(* IEC 61131-3 sources: SortJet_MasterSPS_Aufbau.fbsproj/07_Auftragsverwaltung/BasisSchrittketten (part 2) *)

(* ---- Station_Austransport.fb.st ---- *)
(* METADATA
{
	"v3Meta": {
		"objectGuid": "ceff7ec0-8422-4f2f-902e-5124ad2e42bc"
	}
}
*)
FUNCTION_BLOCK Station_Austransport
VAR_INPUT

  // BOOLEAN
  bpReset                : BOOL;

  // WORD
  wStation               : WORD;
  wWand                  : WORD;

  // STRUKTUR
  Auftragsdaten          : Auftragsdaten_ST;

END_VAR
VAR_OUTPUT

  // BOOLEAN
  bpDone                 : BOOL;
  bpFehler               : BOOL;

END_VAR
VAR

  // BOOLEAN
  blStationQuittiertScheiben      : BOOL;
  blGegenstelleIstShuttle         : BOOL;

  // INT
  ilScheibenZuQuittieren          : INT;

  // WORD
  wlAustransportstation           : WORD;
  wlAustransportstationVorgaenger : WORD;

  // REFERENZ
  Gegenstelle                     : REFERENCE TO StationBasisParameter_ST;

  // STEPS
  steplSchritt           : STEPS_TE;

END_VAR
//-------------------------------------------------------------------------------------------------
// STEUERUNG AUSTRANSPORT
//-------------------------------------------------------------------------------------------------
IF Auftragsdaten.wAuftrag = eStation_Austransport THEN
  CASE steplSchritt OF
    // AUSTRANSPORT =================================
    STEP_0_E:
      (* Hinweis:
         - Ueberpruefung des Sicherheitskreises
      *)
      IF checkSafetyCircuitsNotBlocked(starrStationBasisParameter[wStation], eSKKomponente_Glastransport) THEN
        steplSchritt := STEP_10_E;
      END_IF

    // AUSTRANSPORT ==================================================
    STEP_10_E:
      // ---------------------------------------------------------------------------------------
      //  OPTIONALE - PRUEFUNG DER GLASDATEN
      //
      //  Hinweis:
      // - n/c
      // ---------------------------------------------------------------------------------------
      steplSchritt := STEP_20_E;

      IF NOT AuftragsdatenPruefen( wStation, wWand, Auftragsdaten) THEN
        steplSchritt := STEP_900_E;
      END_IF

    // AUSTRANSPORT =================================
    STEP_20_E:
      (* Hinweis:
         - Uebergabe der Quellstation [Sender] fuer den Austransport [Zum ueberpruefen des Zustandes der Station]
      *)
      wlAustransportstation := Auftragsdaten.wTransferstationsNr1;

      (* Hinweis:
         - Nach einem Systemcheck mit übergroßen Scheiben kann es sein das die Scheibe noch zum Teil auf der Vorgänger Station liegt. Im Systemcheck wird dann "eStation_Warte_Auf_Austransport_Nachfolger" gesetzt
         - Die Station muss dann in Austransport gesetzt weren
      *)

      wlAustransportstationVorgaenger := starrStationBasisParameter[wStation].stMKs.stSchnittstellendaten.wVorgaengerStation;
      IF ( PruefungWertImIntervall( wlAustransportstationVorgaenger, cERSTE_STATION,cLETZTE_STATION ) ) THEN  // Prüfen ob eine gültige Station zugewiesen
        IF ( starrStationBasisParameter[wlAustransportstationVorgaenger].pAuftrag[wWand].wAuftrag = eStation_Warte_Auf_Austransport_Nachfolger ) THEN
          Job_Stationen.AuftragsdatenWand[wlAustransportstationVorgaenger,wWand]         := AuftragsdatenUmkopieren(FALSE, FALSE, Auftragsdaten);
          starrStationBasisParameter[wlAustransportstationVorgaenger].pAuftrag[wWand].wAuftrag := eStation_Austransport;
        END_IF
      END_IF

      (* Hinweis:
         - Zuweisung Transportkopplung
      *)
      CASE wlAustransportstation OF

        // Shuttles
        cERSTES_SHUTTLE..cLETZTES_SHUTTLE:
          (* Hinweis:
             - Transportkopplung
          *)
          IF ( starrStationBasisParameter[wStation].stMKs.stSchnittstellendaten.aAustransporte.Station[Auftragsdaten.wTransferstationsNr1] = Vorwaertig ) THEN
            starrStationBasisParameter[wStation].InGlasTransportNachfolger[wWand] := starrShuttleBasisParameter[Auftragsdaten.wTransferstationsNr1].OutGlasTransport[Auftragsdaten.wTransferwand];
          ELSE
            starrStationBasisParameter[wStation].InGlasTransportVorgaenger[wWand] := starrShuttleBasisParameter[Auftragsdaten.wTransferstationsNr1].OutGlasTransport[Auftragsdaten.wTransferwand];
          END_IF

          steplSchritt := STEP_30_E;

        // Transfershuttles
        //   - Der Auftrag kommt vom TS (TS_Eintransport), hier nur die Transportkopplung
        cERSTES_TRANSFERSHUTTLE..cLETZTES_TRANSFERSHUTTLE:
          IF ( starrStationBasisParameter[wStation].stMKs.stSchnittstellendaten.aAustransporte.Station[Auftragsdaten.wTransferstationsNr1] = Vorwaertig ) THEN
            starrStationBasisParameter[wStation].InGlasTransportNachfolger[wWand] := starrTransfershuttleBasisParameter[Auftragsdaten.wTransferstationsNr1].OutGlasTransport[cWAND_1];
          ELSE
            starrStationBasisParameter[wStation].InGlasTransportVorgaenger[wWand] := starrTransfershuttleBasisParameter[Auftragsdaten.wTransferstationsNr1].OutGlasTransport[cWAND_1];
          END_IF

          steplSchritt := STEP_30_E;

        // Stationen
        cERSTE_STATION..cLETZTE_STATION:

          (* Hinweis:
             - Ist diese Station ein Shuttle, muss sie den Auftrag an die Gegenstelle geben, sofern diese kein Shuttle ist
          *)
          Gegenstelle REF= getBasis( Auftragsdaten.wTransferstationsNr1 );
          blGegenstelleIstShuttle := __ISVALIDREF( Gegenstelle ) AND_THEN __ISVALIDREF( Gegenstelle.stMKs ) AND_THEN Gegenstelle.stMKs.stSchnittstellendaten.bStationIstShuttle;

          // Station ist ein Shuttle
          IF starrStationBasisParameter[wStation].stMKs.stSchnittstellendaten.bStationIstShuttle AND NOT blGegenstelleIstShuttle THEN
            IF ( ( Job_Stationen.AuftragsdatenWand[Auftragsdaten.wTransferstationsNr1, Auftragsdaten.wTransferwand].wAuftrag = eStation_Belegt )
                 OR ( Job_Stationen.AuftragsdatenWand[Auftragsdaten.wTransferstationsNr1, Auftragsdaten.wTransferwand].wAuftrag = eStation_Kein_Auftrag ) )
            THEN

              Job_Stationen.AuftragsdatenWand[Auftragsdaten.wTransferstationsNr1, Auftragsdaten.wTransferwand]          := AuftragsdatenUmkopieren(FALSE, FALSE, Auftragsdaten);
              Job_Stationen.AuftragsdatenWand[Auftragsdaten.wTransferstationsNr1, Auftragsdaten.wTransferwand].wAuftrag := eStation_Eintransport;

              // Transportkopplung
              IF ( starrStationBasisParameter[wStation].stMKs.stSchnittstellendaten.aAustransporte.Station[Auftragsdaten.wTransferstationsNr1] = Vorwaertig ) THEN
                starrStationBasisParameter[wStation].InGlasTransportNachfolger[wWand] := starrStationBasisParameter[Auftragsdaten.wTransferstationsNr1].OutGlasTransport[Auftragsdaten.wTransferwand];
              ELSE
                starrStationBasisParameter[wStation].InGlasTransportVorgaenger[wWand] := starrStationBasisParameter[Auftragsdaten.wTransferstationsNr1].OutGlasTransport[Auftragsdaten.wTransferwand];
              END_IF

              steplSchritt := STEP_30_E;
            END_IF

          ELSE

            // Transportkopplung
            IF ( starrStationBasisParameter[wStation].stMKs.stSchnittstellendaten.aAustransporte.Station[Auftragsdaten.wTransferstationsNr1] = Vorwaertig ) THEN
              starrStationBasisParameter[wStation].InGlasTransportNachfolger[wWand] := starrStationBasisParameter[Auftragsdaten.wTransferstationsNr1].OutGlasTransport[Auftragsdaten.wTransferwand];
            ELSE
              starrStationBasisParameter[wStation].InGlasTransportVorgaenger[wWand] := starrStationBasisParameter[Auftragsdaten.wTransferstationsNr1].OutGlasTransport[Auftragsdaten.wTransferwand];
            END_IF

            steplSchritt := STEP_30_E;

          END_IF

        cERSTE_FREMDANLAGE_AUSLAUF..cLETZTE_FREMDANLAGE_AUSLAUF:
          IF ( Auftragsdaten.wTransferstationsNr2 <> 0 ) THEN
            IF   ( Job_Fremdanlage.AuftragsdatenFremdanlage[wlAustransportstation].wAuftrag = eStation_Kein_Auftrag )
                 AND ( Job_Stationen.AuftragsdatenWand[Auftragsdaten.wTransferstationsNr2, Auftragsdaten.wTransferwand].wAuftrag = eStation_Kein_Auftrag )
            THEN
              steplSchritt := STEP_30_E;
            END_IF
          ELSE
            IF starrStationBasisParameter[wStation].stMKs.stSchnittstellendaten.bStationIstShuttle THEN
              IF ( Job_Fremdanlage.AuftragsdatenFremdanlage[wlAustransportstation].wAuftrag = eStation_Kein_Auftrag ) THEN
                starrStationBasisParameter[wStation].InGlasTransportNachfolger[wWand] := starrFremdanlageAuslaufStationBasisParameter[Auftragsdaten.wTransferstationsNr1].OutGlasTransport[cWAND_1];
                starrFremdanlageAuslaufStationBasisParameter[Auftragsdaten.wTransferstationsNr1].InGlasTransportVorgaenger[cWAND_1] :=  starrStationBasisParameter[wStation].OutGlasTransport[wWand];
                steplSchritt := STEP_30_E;
              END_IF
            ELSE
              starrStationBasisParameter[wStation].InGlasTransportNachfolger[wWand] := starrFremdanlageAuslaufStationBasisParameter[Auftragsdaten.wTransferstationsNr1].OutGlasTransport[cWAND_1];
              starrFremdanlageAuslaufStationBasisParameter[Auftragsdaten.wTransferstationsNr1].InGlasTransportVorgaenger[cWAND_1] :=  starrStationBasisParameter[wStation].OutGlasTransport[wWand];
              steplSchritt := STEP_30_E;
            END_IF
          END_IF

        cERSTE_FREMDANLAGE_EINLAUF..cLETZTE_FREMDANLAGE_EINLAUF:
          ;

        cERSTE_FAECHERWAGENSTATIONS_NR..cLETZTE_FAECHERWAGENSTATIONS_NR:
          ;

        ELSE
          wpgFehlerdaten[0] := starrStationBasisParameter[wStation].stMKs.stStationsNummern.NummerExtern;
          wpgFehlerdaten[1] := wlAustransportstation;
          SpsError( eFehler_Station,
                    cMELDUNG_AUFTRAGSDATEN_FALSCHE_AUSLAUFSTATION,
                    starrStationBasisParameter[wStation].stMKs.stStationsNummern.NummerIntern,
                    AutomatikkreisBestimmen(starrStationBasisParameter[wStation].stMKs.stStationsNummern.NummerSPS),
                    wpgFehlerdaten );

          steplSchritt := STEP_900_E;

      END_CASE

    // AUSTRANSPORT =================================
    STEP_30_E:

      (* Hinweis:
         - Scheibenquittierung
      *)
      ilScheibenZuQuittieren := WORD_TO_INT(Auftragsdaten.wAnzahlScheiben);

      (* Hinweis:
         - Auftragsdaten zuweisen
      *)
      starrStationBasisParameter[wStation].pAuftrag[wWand] := Auftragsdaten;

      (* Hinweis:
         - Auftrags- Optionen bestimmen und zuweisen
      *)
      // Drehen
      starrStationBasisParameter[wStation].pAuftrag[wWand].stAuftragsOptionen.eKippen_SollPosition                  := starrStationBasisParameter[wStation].stMKs.stSchnittstellendaten.aAustransporte.Kippen[Auftragsdaten.wTransferstationsNr1];
      starrStationBasisParameter[wStation].pAuftrag[wWand].stAuftragsOptionen.eKippen_SollPosition_NachEintransport := 0;
      starrStationBasisParameter[wStation].pAuftrag[wWand].stAuftragsOptionen.eKippen_SollPosition_NachAustransport := starrStationBasisParameter[wStation].stMKs.stSchnittstellendaten.aAustransporte.KippenNachAustransport[Auftragsdaten.wTransferstationsNr1];

      IF ( Auftragsdaten.rAuftragsDicke < wgUnterteilerMinMaxGlasdicke ) THEN
        starrStationBasisParameter[wStation].pAuftrag[wWand].stAuftragsOptionen.eDickenverstellung := eZylinderStellung16mm;
      ELSE
        starrStationBasisParameter[wStation].pAuftrag[wWand].stAuftragsOptionen.eDickenverstellung := eZylinderStellung29mm;
      END_IF
      IF starrStationBasisParameter[wStation].stMKs.stStationsOptionen.stDrehstation.bDrehpositionenVomMMI THEN
        starrStationBasisParameter[wStation].pAuftrag[wWand].stAuftragsOptionen.eDrehen_Sollposition                 := REAL_TO_WORD(Auftragsdaten.rStationsZielposition);
        starrStationBasisParameter[wStation].pAuftrag[wWand].stAuftragsOptionen.eDrehen_Sollposition_NachAustransport := REAL_TO_WORD(Auftragsdaten.rTransferposition2);
      ELSE
        starrStationBasisParameter[wStation].pAuftrag[wWand].stAuftragsOptionen.eDrehen_Sollposition                 := starrStationBasisParameter[wStation].stMKs.stSchnittstellendaten.aAustransporte.Drehen[Auftragsdaten.wTransferstationsNr1];
        starrStationBasisParameter[wStation].pAuftrag[wWand].stAuftragsOptionen.eDrehen_Sollposition_NachAustransport := starrStationBasisParameter[wStation].stMKs.stSchnittstellendaten.aAustransporte.DrehenNachAustransport[Auftragsdaten.wTransferstationsNr1];
      END_IF
      starrStationBasisParameter[wStation].pAuftrag[wWand].stAuftragsOptionen.eDrehen_Sollposition_NachEintransport := 0;
      starrStationBasisParameter[wStation].pAuftrag[wWand].stAuftragsOptionen.eGlastransport := starrStationBasisParameter[wStation].stMKs.stSchnittstellendaten.aAustransporte.Glastransport[Auftragsdaten.wTransferstationsNr1];
      starrStationBasisParameter[wStation].pAuftrag[wWand].stAuftragsOptionen.eHub                  := starrStationBasisParameter[wStation].stMKs.stSchnittstellendaten.aAustransporte.Hub[Auftragsdaten.wTransferstationsNr1];
      starrStationBasisParameter[wStation].pAuftrag[wWand].stAuftragsOptionen.eHub_NachEintransport := 0;
      starrStationBasisParameter[wStation].pAuftrag[wWand].stAuftragsOptionen.eHub_NachAustransport := starrStationBasisParameter[wStation].stMKs.stSchnittstellendaten.aAustransporte.HubNachAustransport[Auftragsdaten.wTransferstationsNr1];
      starrStationBasisParameter[wStation].pAuftrag[wWand].stAuftragsOptionen.eQuerachse := 0;
      starrStationBasisParameter[wStation].pAuftrag[wWand].stAuftragsOptionen.eAchsrichtung := starrStationBasisParameter[wStation].stMKs.stSchnittstellendaten.aAustransporte.Achsrichtung[Auftragsdaten.wTransferstationsNr1];
      starrStationBasisParameter[wStation].pAuftrag[wWand].stAuftragsOptionen.wMaxTransportGeschwindigkeit:= 0;

      starrStationBasisParameter[wStation].bScheibentrennen[wWand] := FALSE;
      starrStationBasisParameter[wStation].bRueckwaertsTransportieren[wWand] := ( starrStationBasisParameter[wStation].stMKs.stSchnittstellendaten.aAustransporte.Station[Auftragsdaten.wTransferstationsNr1] = Rueckwaertig );

      steplSchritt := STEP_35_E;

    // AUSTRANSPORT =================================
    STEP_35_E:
      // Im Step 35 wird in dem vererbten FB Anlagenspezifische Auftragsoptionen gesetzt
      starrStationBasisParameter[wStation].bAustransport[wWand] := TRUE;
      steplSchritt := STEP_40_E;

    // AUSTRANSPORT =================================
    STEP_40_E:

      (* Hinweis:
         - Scheibenzaehler dekrementieren
         - Scheibe quittieren, sofern dies nötig ist
      *)
      blStationQuittiertScheiben := starrStationBasisParameter[wStation].stMKs.stSchnittstellendaten.aAustransporte.bStationQuittiertScheibe[wlAustransportstation];

      IF ( starrStationBasisParameter[wStation].OutGlasTransport[wWand].bQuittScheibe ) THEN

        IF ( ilScheibenZuQuittieren > 0 ) AND blStationQuittiertScheiben THEN

          wSps2MmiZielStation  := Auftragsdaten.wTransferstationsNr1;
          wSps2MmiQuellStation := starrStationBasisParameter[wStation].stMKs.stStationsNummern.NummerIntern;
          wSps2MmiZielWand     := Auftragsdaten.wTransferwand;
          wSps2MmiQuellWand    := Auftragsdaten.wStationsWand;
          dwSps2MmiWartezeit   := starrStationBasisParameter[wStation].dwWartezeit[wWand];

          IF starrStationBasisParameter[wStation].stMKs.stSchnittstellendaten.bStationIstShuttle THEN
            wSPS2MMIAuftragstyp  := 1;
          ELSE
            wSPS2MMIAuftragstyp  := 0;
          END_IF;

          MsgToMmi(auftragsnr_w := SB0_SPS_QUIT_SHEET_ORDER );

        END_IF

        ilScheibenZuQuittieren := ilScheibenZuQuittieren - 1;

      END_IF

      (* Hinweis:
         - Abschliessen des Austransport
      *)
      IF ( starrStationBasisParameter[wStation].bAustransportAbgeschlossen[wWand] ) THEN
        starrStationBasisParameter[wStation].bRueckwaertsTransportieren[wWand] := FALSE;
        starrStationBasisParameter[wStation].bAustransport[wWand] := FALSE;
        steplSchritt := STEP_100_E;
      END_IF

      (* Fehlerbehandlung:
         - Station
      *)
      IF ( starrStationBasisParameter[wStation].bFehler ) THEN
        SpsError( eFehler_Station,
                  starrStationBasisParameter[wStation].wFehlerNummer,
                  starrStationBasisParameter[wStation].stMKs.stStationsNummern.NummerIntern,
                  AutomatikkreisBestimmen(starrStationBasisParameter[wStation].stMKs.stStationsNummern.NummerSPS),
                  starrStationBasisParameter[wStation].awFehlerInformationen );

        starrStationBasisParameter[wStation].bAustransport[wWand] := FALSE;
        starrStationBasisParameter[wStation].bRueckwaertsTransportieren[wWand] := FALSE;
        steplSchritt := STEP_900_E;
      END_IF

    // AUSTRANSPORT ==============================================
    STEP_100_E:
      (* Anmerkung:
         - Gueltige Anzahl von Scheiben wurden quittiert
      *)
      IF ( ilScheibenZuQuittieren = 0 ) THEN
        steplSchritt := STEP_1000_E;

      (* Anmerkung:
         - Zu wenig Scheiben quittiert
      *)
      ELSIF ( ilScheibenZuQuittieren > 0 ) THEN
        wpgFehlerdaten[0] := starrStationBasisParameter[wStation].stMKs.stStationsNummern.NummerExtern;
        wpgFehlerdaten[1] := wWand;

        SpsError( eFehler_Station,
                  cMELDUNG_STATION_ZUWENIG_SCHEIBEN_QUITTIERT_AUSTRANSPORT,
                  starrStationBasisParameter[wStation].stMKs.stStationsNummern.NummerIntern,
                  AutomatikkreisBestimmen(starrStationBasisParameter[wStation].stMKs.stStationsNummern.NummerSPS),
                  wpgFehlerdaten );

        steplSchritt := STEP_900_E;

      (* Anmerkung:
         - Zu viele Scheiben quittiert
      *)
      ELSIF ( ilScheibenZuQuittieren < 0 ) THEN
        wpgFehlerdaten[0] := starrStationBasisParameter[wStation].stMKs.stStationsNummern.NummerExtern;
        wpgFehlerdaten[1] := wWand;

        SpsError( eFehler_Station,
                  cMELDUNG_STATION_ZUVIELE_SCHEIBEN_QUITTIERT_AUSTRANSPORT,
                  starrStationBasisParameter[wStation].stMKs.stStationsNummern.NummerIntern,
                  AutomatikkreisBestimmen(starrStationBasisParameter[wStation].stMKs.stStationsNummern.NummerSPS),
                  wpgFehlerdaten );

        steplSchritt := STEP_900_E;
      END_IF

    // AUSTRANSPORT =================================
    STEP_900_E:
      bpFehler := TRUE;

    // AUSTRANSPORT =================================
    STEP_1000_E:
      bpDone := TRUE;
      IF Auftragsdaten.stAuftragsInformationen.cBIT_SRCSTATION_EMPTY THEN
        Auftragsdaten.wAuftrag := eStation_Kein_Auftrag;
      ELSE
        Auftragsdaten.wAuftrag := eStation_Belegt;
      END_IF
  END_CASE

END_IF

IF bpReset THEN
  bpFehler := FALSE;
  bpReset := FALSE;
  bpDone := FALSE;
  steplSchritt := STEP_0_E;
  starrStationBasisParameter[wStation].bRueckwaertsTransportieren[wWand] := FALSE;
  starrStationBasisParameter[wStation].bAustransport[wWand] := FALSE;
END_IF
END_FUNCTION_BLOCK

(* ---- Station_Durchtransport.fb.st ---- *)
(* METADATA
{
	"v3Meta": {
		"objectGuid": "2b51cd18-a11d-48d6-a685-bb5f301afb70"
	}
}
*)
FUNCTION_BLOCK Station_Durchtransport
VAR_INPUT

  // BOOLEAN
  bpReset                : BOOL;

  // WORD
  wStation               : WORD;
  wWand                  : WORD;

  // STRUKTUR
  Auftragsdaten          : Auftragsdaten_ST;

END_VAR
VAR_OUTPUT

  // BOOLEAN
  bpDone                 : BOOL;
  bpFehler               : BOOL;

END_VAR
VAR

  // BOOLEAN
  blStationQuittiertScheiben             : BOOL;
  blKopplungGefundenEintransport         : BOOL;
  blKopplungGefundenAustransport         : BOOL;

  // INT
  ilScheibenZuQuittieren : INT;

  // WORD
  wlEintransportstation : WORD;
  wlAustransportstation : WORD;

  // STEPS
  steplSchritt           : STEPS_TE;

END_VAR
//-------------------------------------------------------------------------------------------------
// STEUERUNG DURCHTRANSPORT
//-------------------------------------------------------------------------------------------------
IF Auftragsdaten.wAuftrag = eStation_Durchtransport THEN
  CASE steplSchritt OF
    // DURCHTRANSPORT =================================
    STEP_0_E:
      (* Hinweis:
         - Ueberpruefung des Sicherheitskreises
      *)
      IF checkSafetyCircuitsNotBlocked(starrStationBasisParameter[wStation], eSKKomponente_Glastransport) THEN
        steplSchritt := STEP_10_E;
      END_IF

    // DURCHTRANSPORT ==================================================
    STEP_10_E:
      // ---------------------------------------------------------------------------------------
      //  OPTIONALE - PRUEFUNG DER GLASDATEN
      //
      //  Hinweis:
      // - n/c
      // ---------------------------------------------------------------------------------------
      steplSchritt := STEP_20_E;

      IF NOT AuftragsdatenPruefen( wStation, wWand, Auftragsdaten) THEN
        steplSchritt := STEP_900_E;
      END_IF

    // DURCHTRANSPORT =================================
    STEP_20_E:
      (* Hinweis:
         - Kopplung fuer diesen Auftrag neu bestimmen. Sonst ueberschreibt ein Merker aus dem letzten Auftrag den Fehlerschritt.
      *)
      blKopplungGefundenEintransport := FALSE;
      blKopplungGefundenAustransport := FALSE;

      (* Hinweis:
         - Uebergabe der Quellstation [Sender] fuer den Austransport [Zum ueberpruefen des Zustandes der Station]
      *)
      wlEintransportstation := Auftragsdaten.wTransferstationsNr1;
      wlAustransportstation := Auftragsdaten.wTransferstationsNr2;

      (* Hinweis:
         - Zuweisung Transportkopplung
      *)
      CASE wlEintransportstation OF

        // Shuttles
        cERSTES_SHUTTLE..cLETZTES_SHUTTLE:
          (* Hinweis:
             - Transportkopplung
          *)
          IF ( starrStationBasisParameter[wStation].stMKs.stSchnittstellendaten.aEintransporte.Station[wlEintransportstation] = Vorwaertig ) THEN
            starrStationBasisParameter[wStation].InGlasTransportVorgaenger[wWand] := starrShuttleBasisParameter[wlEintransportstation].OutGlasTransport[Auftragsdaten.wTransferwand];
          ELSE
            starrStationBasisParameter[wStation].InGlasTransportNachfolger[wWand] := starrShuttleBasisParameter[wlEintransportstation].OutGlasTransport[Auftragsdaten.wTransferwand];
          END_IF
          blKopplungGefundenEintransport := TRUE;

        // Stationen
        cERSTE_STATION..cLETZTE_STATION:
          (* Hinweis:
             - Transportkopplung
          *)
          IF ( starrStationBasisParameter[wStation].stMKs.stSchnittstellendaten.aEintransporte.Station[wlEintransportstation] = Vorwaertig ) THEN
            starrStationBasisParameter[wStation].InGlasTransportVorgaenger[wWand] := starrStationBasisParameter[wlEintransportstation].OutGlasTransport[Auftragsdaten.wTransferwand];
          ELSE
            starrStationBasisParameter[wStation].InGlasTransportNachfolger[wWand] := starrStationBasisParameter[wlEintransportstation].OutGlasTransport[Auftragsdaten.wTransferwand];
          END_IF
          blKopplungGefundenEintransport := TRUE;

        cERSTE_FREMDANLAGE_AUSLAUF..cLETZTE_FREMDANLAGE_AUSLAUF:
          (* Hinweis:
             - Transportkopplung
          *)
          IF ( starrStationBasisParameter[wStation].stMKs.stSchnittstellendaten.aEintransporte.Station[wlEintransportstation] = Vorwaertig ) THEN
            starrStationBasisParameter[wStation].InGlasTransportVorgaenger[wWand] := starrFremdanlageAuslaufStationBasisParameter[wlEintransportstation].OutGlasTransport[cWAND_1];
          ELSE
            starrStationBasisParameter[wStation].InGlasTransportNachfolger[wWand] := starrFremdanlageAuslaufStationBasisParameter[wlEintransportstation].OutGlasTransport[cWAND_1];
          END_IF
          blKopplungGefundenEintransport := TRUE;

        ELSE
          wpgFehlerdaten[0] := starrStationBasisParameter[wStation].stMKs.stStationsNummern.NummerExtern;
          wpgFehlerdaten[1] := wlEintransportstation;
          SpsError( eFehler_Station,
                    cMELDUNG_AUFTRAGSDATEN_FALSCHE_EINLAUFSTATION,
                    starrStationBasisParameter[wStation].stMKs.stStationsNummern.NummerIntern,
                    AutomatikkreisBestimmen(starrStationBasisParameter[wStation].stMKs.stStationsNummern.NummerSPS),
                    wpgFehlerdaten );

          steplSchritt := STEP_900_E;

      END_CASE

      (* Hinweis:
         - Zuweisung Transportkopplung
      *)
      CASE wlAustransportstation OF

        // Shuttles
        cERSTES_SHUTTLE..cLETZTES_SHUTTLE:
          (* Hinweis:
             - Transportkopplung
          *)
          IF ( starrStationBasisParameter[wStation].stMKs.stSchnittstellendaten.aAustransporte.Station[wlAustransportstation] = Vorwaertig ) THEN
            starrStationBasisParameter[wStation].InGlasTransportNachfolger[wWand] := starrShuttleBasisParameter[wlAustransportstation].OutGlasTransport[Auftragsdaten.wTransferwand];
          ELSE
            starrStationBasisParameter[wStation].InGlasTransportVorgaenger[wWand] := starrShuttleBasisParameter[wlAustransportstation].OutGlasTransport[Auftragsdaten.wTransferwand];
          END_IF
          blKopplungGefundenAustransport := TRUE;

        // Stationen
        cERSTE_STATION..cLETZTE_STATION:
          (* Hinweis:
             - Transportkopplung
          *)
          IF ( starrStationBasisParameter[wStation].stMKs.stSchnittstellendaten.aAustransporte.Station[wlAustransportstation] = Vorwaertig ) THEN
            starrStationBasisParameter[wStation].InGlasTransportNachfolger[wWand] := starrStationBasisParameter[wlAustransportstation].OutGlasTransport[Auftragsdaten.wTransferwand];
          ELSE
            starrStationBasisParameter[wStation].InGlasTransportVorgaenger[wWand] := starrStationBasisParameter[wlAustransportstation].OutGlasTransport[Auftragsdaten.wTransferwand];
          END_IF
          blKopplungGefundenAustransport := TRUE;

        cERSTE_FREMDANLAGE_AUSLAUF..cLETZTE_FREMDANLAGE_AUSLAUF:
          (* Hinweis:
             - Transportkopplung
          *)
          IF ( starrStationBasisParameter[wStation].stMKs.stSchnittstellendaten.aAustransporte.Station[wlAustransportstation] = Vorwaertig ) THEN
            starrStationBasisParameter[wStation].InGlasTransportNachfolger[wWand] := starrFremdanlageAuslaufStationBasisParameter[wlAustransportstation].OutGlasTransport[cWAND_1];
          ELSE
            starrStationBasisParameter[wStation].InGlasTransportVorgaenger[wWand] := starrFremdanlageAuslaufStationBasisParameter[wlAustransportstation].OutGlasTransport[cWAND_1];
          END_IF
          blKopplungGefundenAustransport := TRUE;

        ELSE
          wpgFehlerdaten[0] := starrStationBasisParameter[wStation].stMKs.stStationsNummern.NummerExtern;
          wpgFehlerdaten[1] := wlAustransportstation;
          SpsError( eFehler_Station,
                    cMELDUNG_AUFTRAGSDATEN_FALSCHE_AUSLAUFSTATION,
                    starrStationBasisParameter[wStation].stMKs.stStationsNummern.NummerIntern,
                    AutomatikkreisBestimmen(starrStationBasisParameter[wStation].stMKs.stStationsNummern.NummerSPS),
                    wpgFehlerdaten );

          steplSchritt := STEP_900_E;

      END_CASE

      IF blKopplungGefundenEintransport AND blKopplungGefundenAustransport THEN
        steplSchritt := STEP_30_E;
      END_IF

    // DURCHTRANSPORT =================================
    STEP_30_E:

      (* Hinweis:
         - Scheibenquittierung
      *)
      ilScheibenZuQuittieren := WORD_TO_INT(Auftragsdaten.wAnzahlScheiben);

      (* Hinweis:
         - Auftragsdaten zuweisen
      *)
      starrStationBasisParameter[wStation].pAuftrag[wWand] := Auftragsdaten;

      (* Hinweis:
         - Auftrags- Optionen bestimmen und zuweisen
      *)
      starrStationBasisParameter[wStation].pAuftrag[wWand].stAuftragsOptionen.eKippen_SollPosition := starrStationBasisParameter[wStation].stMKs.stSchnittstellendaten.aEintransporte.Kippen[wlEintransportstation];

      IF ( Auftragsdaten.rAuftragsDicke < wgUnterteilerMinMaxGlasdicke ) THEN
        starrStationBasisParameter[wStation].pAuftrag[wWand].stAuftragsOptionen.eDickenverstellung := eZylinderStellung16mm;
      ELSE
        starrStationBasisParameter[wStation].pAuftrag[wWand].stAuftragsOptionen.eDickenverstellung := eZylinderStellung29mm;
      END_IF
      starrStationBasisParameter[wStation].pAuftrag[wWand].stAuftragsOptionen.eDrehen_Sollposition := 0;
      starrStationBasisParameter[wStation].pAuftrag[wWand].stAuftragsOptionen.eDrehen_Sollposition_NachAustransport := 0;
      starrStationBasisParameter[wStation].pAuftrag[wWand].stAuftragsOptionen.eKippen_SollPosition_NachAustransport := 0;
      starrStationBasisParameter[wStation].pAuftrag[wWand].stAuftragsOptionen.eGlastransport := starrStationBasisParameter[wStation].stMKs.stSchnittstellendaten.aEintransporte.Glastransport[wlEintransportstation];
      starrStationBasisParameter[wStation].pAuftrag[wWand].stAuftragsOptionen.eHub                  := starrStationBasisParameter[wStation].stMKs.stSchnittstellendaten.aEintransporte.Hub[wlEintransportstation];
      starrStationBasisParameter[wStation].pAuftrag[wWand].stAuftragsOptionen.eHub_NachEintransport := 0;
      starrStationBasisParameter[wStation].pAuftrag[wWand].stAuftragsOptionen.eHub_NachAustransport := 0;
      starrStationBasisParameter[wStation].pAuftrag[wWand].stAuftragsOptionen.eQuerachse := 0;
      starrStationBasisParameter[wStation].pAuftrag[wWand].stAuftragsOptionen.eAchsrichtung := 0;
      starrStationBasisParameter[wStation].pAuftrag[wWand].stAuftragsOptionen.wMaxTransportGeschwindigkeit:= 0;
      starrStationBasisParameter[wStation].pAuftrag[wWand].stAuftragsOptionen.eDrehen_Sollposition_NachEintransport := 0;
      starrStationBasisParameter[wStation].pAuftrag[wWand].stAuftragsOptionen.eKippen_SollPosition_NachEintransport := 0;

      starrStationBasisParameter[wStation].bScheibentrennen[wWand]           := FALSE;
      starrStationBasisParameter[wStation].bRueckwaertsTransportieren[wWand] := ( starrStationBasisParameter[wStation].stMKs.stSchnittstellendaten.aEintransporte.Station[wlEintransportstation] = Rueckwaertig )
                                                                                AND ( starrStationBasisParameter[wStation].stMKs.stSchnittstellendaten.aAustransporte.Station[wlAustransportstation] = Rueckwaertig );
      starrStationBasisParameter[wStation].bDurchtransport[wWand]            := TRUE;

      steplSchritt := STEP_40_E;

    // AUSTRANSPORT =================================
    STEP_40_E:

      (* Hinweis:
         - Scheibenzaehler dekrementieren
         - Scheibe quittieren, sofern dies nötig ist
      *)
      blStationQuittiertScheiben := TRUE;

      IF ( starrStationBasisParameter[wStation].OutGlasTransport[wWand].bQuittScheibe ) THEN

        IF ( ilScheibenZuQuittieren > 0 ) AND blStationQuittiertScheiben THEN

          wSps2MmiZielStation  := starrStationBasisParameter[wStation].stMKs.stStationsNummern.NummerIntern;
          wSps2MmiQuellStation := wlEintransportstation;
          wSps2MmiZielWand     := Auftragsdaten.wStationsWand;
          wSps2MmiQuellWand    := Auftragsdaten.wTransferwand;
          dwSps2MmiWartezeit   := starrStationBasisParameter[wStation].dwWartezeit[wWand];
          wSPS2MMIAuftragstyp  := 0;

          MsgToMmi(auftragsnr_w := SB0_SPS_QUIT_SHEET_ORDER );

        END_IF

        ilScheibenZuQuittieren := ilScheibenZuQuittieren - 1;

      END_IF

      (* Hinweis:
         - Abschliessen des Austransport
      *)
      IF ( starrStationBasisParameter[wStation].bDurchtransportAbgeschlossen[wWand] ) THEN
        starrStationBasisParameter[wStation].bRueckwaertsTransportieren[wWand] := FALSE;
        starrStationBasisParameter[wStation].bDurchtransport[wWand] := FALSE;
        steplSchritt := STEP_1000_E;
      END_IF

      (* Fehlerbehandlung:
         - Station
      *)
      IF ( starrStationBasisParameter[wStation].bFehler ) THEN
        SpsError( eFehler_Station,
                  starrStationBasisParameter[wStation].wFehlerNummer,
                  starrStationBasisParameter[wStation].stMKs.stStationsNummern.NummerIntern,
                  AutomatikkreisBestimmen(starrStationBasisParameter[wStation].stMKs.stStationsNummern.NummerSPS),
                  starrStationBasisParameter[wStation].awFehlerInformationen );
        starrStationBasisParameter[wStation].bDurchtransport[wWand] := FALSE;
        starrStationBasisParameter[wStation].bRueckwaertsTransportieren[wWand] := FALSE;
        steplSchritt := STEP_900_E;
      END_IF

    // DURCHTRANSPORT =================================
    STEP_900_E:
      bpFehler := TRUE;

    // DURCHTRANSPORT =================================
    STEP_1000_E:
      bpDone := TRUE;
      Auftragsdaten.wAuftrag := eStation_Kein_Auftrag;

  END_CASE

END_IF

IF bpReset THEN
  bpFehler := FALSE;
  bpReset := FALSE;
  bpDone := FALSE;
  blKopplungGefundenEintransport := FALSE;
  blKopplungGefundenAustransport := FALSE;
  blStationQuittiertScheiben := FALSE;
  steplSchritt := STEP_0_E;
  starrStationBasisParameter[wStation].bRueckwaertsTransportieren[wWand] := FALSE;
  starrStationBasisParameter[wStation].bDurchtransport[wWand] := FALSE;
END_IF
END_FUNCTION_BLOCK

(* ---- Station_Eintransport.fb.st ---- *)
(* METADATA
{
	"v3Meta": {
		"objectGuid": "db6c6d03-f822-435f-8f93-f5a504a5ce8d"
	}
}
*)
FUNCTION_BLOCK Station_Eintransport
VAR_INPUT

  // BOOLEAN
  bpReset                : BOOL;

  // WORD
  wStation               : WORD;
  wWand                  : WORD;

  // STRUKTUR
  Auftragsdaten          : Auftragsdaten_ST;

END_VAR
VAR_OUTPUT

  // BOOLEAN
  bpDone                 : BOOL;
  bpFehler               : BOOL;

END_VAR
VAR

  // BOOLEAN
  blStationQuittiertScheiben : BOOL;
  blGegenstelleIstShuttle    : BOOL;

  // WORD
  wlEintransportstation  : WORD;

  // INT
  ilScheibenZuQuittieren : INT;

  // REFERENZ
  Gegenstelle            : REFERENCE TO StationBasisParameter_ST;

  // STEPS
  steplSchritt           : STEPS_TE;

END_VAR
//-------------------------------------------------------------------------------------------------
// STEUERUNG: EINTRANSPORT
//-------------------------------------------------------------------------------------------------
IF ( Auftragsdaten.wAuftrag = eStation_Eintransport ) THEN
  CASE steplSchritt OF
    // EINTRANSPORT ==================================================
    STEP_0_E:
      (* Hinweis:
         - Ueberpruefung des Sicherheitskreises
      *)
      IF checkSafetyCircuitsNotBlocked(starrStationBasisParameter[wStation], eSKKomponente_Glastransport) THEN
        steplSchritt := STEP_10_E;
      END_IF

    // EINTRANSPORT ==================================================
    STEP_10_E:
      // ---------------------------------------------------------------------------------------
      //  OPTIONALE - PRUEFUNG DER GLASDATEN
      //
      //  Hinweis:
      // - n/c
      // ---------------------------------------------------------------------------------------
      steplSchritt := STEP_20_E;

      IF NOT AuftragsdatenPruefen( wStation, wWand, Auftragsdaten) THEN
        steplSchritt := STEP_900_E;
      END_IF

    // EINTRANSPORT ==================================================
    STEP_20_E:
      // ---------------------------------------------------------------------------------------
      //  OPTIONALE - PRUEFUNG DER GLASDATEN
      //
      //  Hinweis:
      // - n/c
      // ---------------------------------------------------------------------------------------

      // Glastyp festlegen
      IF ( Auftragsdaten.rAuftragsLaenge > starrStationBasisParameter[wStation].stMKs.stStationsParameter.rLaengeUebergroesseScheibe ) THEN
        starrStationBasisParameter[wStation].wGlasTyp[wWand] := eScheibe_Maximal;
      ELSE
        starrStationBasisParameter[wStation].wGlasTyp[wWand] := eScheibe_Default;
      END_IF

      steplSchritt := STEP_30_E;

    // EINTRANSPORT ==================================================
    STEP_30_E:
      (* Hinweis:
         - Uebergabe der Quellstation [Sender] fuer den Austransport [Zum ueberpruefen des Zustandes der Station]
      *)
      wlEintransportstation := Auftragsdaten.wTransferstationsNr1;

      (* Hinweis:
         - Zuweisung Transportkopplung
      *)
      CASE wlEintransportstation OF

        // Shuttles
        cERSTES_SHUTTLE..cLETZTES_SHUTTLE:
          (* Hinweis:
             - Transportkopplung
          *)
          IF ( starrStationBasisParameter[wStation].stMKs.stSchnittstellendaten.aEintransporte.Station[Auftragsdaten.wTransferstationsNr1] = Vorwaertig ) THEN
            starrStationBasisParameter[wStation].InGlasTransportVorgaenger[wWand] := starrShuttleBasisParameter[Auftragsdaten.wTransferstationsNr1].OutGlasTransport[Auftragsdaten.wTransferwand];
          ELSE
            starrStationBasisParameter[wStation].InGlasTransportNachfolger[wWand] := starrShuttleBasisParameter[Auftragsdaten.wTransferstationsNr1].OutGlasTransport[Auftragsdaten.wTransferwand];
          END_IF

          steplSchritt := STEP_40_E;

        // Transfershuttles
        //   - Der Auftrag kommt vom TS (TS_Austransport), hier nur die Transportkopplung
        cERSTES_TRANSFERSHUTTLE..cLETZTES_TRANSFERSHUTTLE:
          IF ( starrStationBasisParameter[wStation].stMKs.stSchnittstellendaten.aEintransporte.Station[Auftragsdaten.wTransferstationsNr1] = Vorwaertig ) THEN
            starrStationBasisParameter[wStation].InGlasTransportVorgaenger[wWand] := starrTransfershuttleBasisParameter[Auftragsdaten.wTransferstationsNr1].OutGlasTransport[cWAND_1];
          ELSE
            starrStationBasisParameter[wStation].InGlasTransportNachfolger[wWand] := starrTransfershuttleBasisParameter[Auftragsdaten.wTransferstationsNr1].OutGlasTransport[cWAND_1];
          END_IF

          steplSchritt := STEP_40_E;

        // Stationen
        cERSTE_STATION..cLETZTE_STATION:

          (* Hinweis:
             - Ist die Gegenstelle selbst ein Shuttle, bekommt sie keinen Auftrag von uns, wir bekommen ihn von ihr
          *)
          Gegenstelle REF= getBasis( wlEintransportstation );
          blGegenstelleIstShuttle := __ISVALIDREF( Gegenstelle ) AND_THEN __ISVALIDREF( Gegenstelle.stMKs ) AND_THEN Gegenstelle.stMKs.stSchnittstellendaten.bStationIstShuttle;

          IF ( ( Job_Stationen.AuftragsdatenWand[Auftragsdaten.wTransferstationsNr1, Auftragsdaten.wTransferwand].wAuftrag = eStation_Belegt )
               OR ( Job_Stationen.AuftragsdatenWand[Auftragsdaten.wTransferstationsNr1, Auftragsdaten.wTransferwand].wAuftrag = eStation_Warte_Auf_Austransport ) )
             OR blGegenstelleIstShuttle
          THEN

            // Ist der Vorgänger ein Shuttle, dann keinen Auftrag schreiben... Wir kriegen dann den Auftrag von ihm
            IF NOT blGegenstelleIstShuttle THEN
              Job_Stationen.AuftragsdatenWand[Auftragsdaten.wTransferstationsNr1, Auftragsdaten.wTransferwand]          := AuftragsdatenUmkopieren(FALSE, FALSE, Auftragsdaten);
              Job_Stationen.AuftragsdatenWand[Auftragsdaten.wTransferstationsNr1, Auftragsdaten.wTransferwand].wAuftrag := eStation_Austransport;
            END_IF

            // Transportkopplung
            IF ( starrStationBasisParameter[wStation].stMKs.stSchnittstellendaten.aEintransporte.Station[Auftragsdaten.wTransferstationsNr1] = Vorwaertig ) THEN
              starrStationBasisParameter[wStation].InGlasTransportVorgaenger[wWand] := starrStationBasisParameter[Auftragsdaten.wTransferstationsNr1].OutGlasTransport[Auftragsdaten.wTransferwand];
            ELSE
              starrStationBasisParameter[wStation].InGlasTransportNachfolger[wWand] := starrStationBasisParameter[Auftragsdaten.wTransferstationsNr1].OutGlasTransport[Auftragsdaten.wTransferwand];
            END_IF

            steplSchritt := STEP_40_E;
          END_IF

        cERSTE_FREMDANLAGE_AUSLAUF..cLETZTE_FREMDANLAGE_AUSLAUF:
          ;

        cERSTE_FREMDANLAGE_EINLAUF..cLETZTE_FREMDANLAGE_EINLAUF:
          ;

        cERSTE_FAECHERWAGENSTATIONS_NR..cLETZTE_FAECHERWAGENSTATIONS_NR:
          ;

        ELSE
          wpgFehlerdaten[0] := starrStationBasisParameter[wStation].stMKs.stStationsNummern.NummerExtern;
          wpgFehlerdaten[1] := wlEintransportstation;
          SpsError( eFehler_Station,
                    cMELDUNG_AUFTRAGSDATEN_FALSCHE_EINLAUFSTATION,
                    starrStationBasisParameter[wStation].stMKs.stStationsNummern.NummerIntern,
                    AutomatikkreisBestimmen(starrStationBasisParameter[wStation].stMKs.stStationsNummern.NummerSPS),
                    wpgFehlerdaten );

          steplSchritt := STEP_900_E;

      END_CASE

    // EINTRANSPORT ==================================================
    STEP_40_E:
      (* Hinweis:
         - Scheibenquittierung
      *)
      ilScheibenZuQuittieren := WORD_TO_INT(Auftragsdaten.wAnzahlScheiben);

      (* Hinweis:
         - Auftragsdaten zuweisen
      *)
      starrStationBasisParameter[wStation].pAuftrag[wWand] := Auftragsdaten;

      (* Hinweis:
         - Auftrags- Optionen bestimmen und zuweisen
      *)
      // Kippen
      starrStationBasisParameter[wStation].pAuftrag[wWand].stAuftragsOptionen.eKippen_SollPosition                  := starrStationBasisParameter[wStation].stMKs.stSchnittstellendaten.aEintransporte.Kippen[Auftragsdaten.wTransferstationsNr1];
      starrStationBasisParameter[wStation].pAuftrag[wWand].stAuftragsOptionen.eKippen_SollPosition_NachEintransport := starrStationBasisParameter[wStation].stMKs.stSchnittstellendaten.aEintransporte.KippenNachEintransport[Auftragsdaten.wTransferstationsNr1];
      starrStationBasisParameter[wStation].pAuftrag[wWand].stAuftragsOptionen.eKippen_SollPosition_NachAustransport := 0;

      IF ( Auftragsdaten.rAuftragsDicke < wgMKScheibenDicke13mm ) THEN
        starrStationBasisParameter[wStation].pAuftrag[wWand].stAuftragsOptionen.eDickenverstellung := eZylinderStellung16mm;
      ELSIF ( Auftragsdaten.rAuftragsDicke <= wgMKScheibenDicke19mm ) THEN
        starrStationBasisParameter[wStation].pAuftrag[wWand].stAuftragsOptionen.eDickenverstellung := eZylinderStellung23mm;
      ELSE
        starrStationBasisParameter[wStation].pAuftrag[wWand].stAuftragsOptionen.eDickenverstellung := eZylinderStellung29mm;
      END_IF

      IF starrStationBasisParameter[wStation].stMKs.stStationsOptionen.stDrehstation.bDrehpositionenVomMMI THEN
        starrStationBasisParameter[wStation].pAuftrag[wWand].stAuftragsOptionen.eDrehen_Sollposition                 := REAL_TO_WORD(Auftragsdaten.rStationsZielposition);
        starrStationBasisParameter[wStation].pAuftrag[wWand].stAuftragsOptionen.eDrehen_Sollposition_NachEintransport := REAL_TO_WORD(Auftragsdaten.rTransferposition2);
      ELSE
        starrStationBasisParameter[wStation].pAuftrag[wWand].stAuftragsOptionen.eDrehen_Sollposition                 := starrStationBasisParameter[wStation].stMKs.stSchnittstellendaten.aEintransporte.Drehen[Auftragsdaten.wTransferstationsNr1];
        starrStationBasisParameter[wStation].pAuftrag[wWand].stAuftragsOptionen.eDrehen_Sollposition_NachEintransport := starrStationBasisParameter[wStation].stMKs.stSchnittstellendaten.aEintransporte.DrehenNachEintransport[Auftragsdaten.wTransferstationsNr1];
      END_IF
      starrStationBasisParameter[wStation].pAuftrag[wWand].stAuftragsOptionen.eDrehen_Sollposition_NachAustransport := 0;
      starrStationBasisParameter[wStation].pAuftrag[wWand].stAuftragsOptionen.eGlastransport := starrStationBasisParameter[wStation].stMKs.stSchnittstellendaten.aEintransporte.Glastransport[Auftragsdaten.wTransferstationsNr1];
      starrStationBasisParameter[wStation].pAuftrag[wWand].stAuftragsOptionen.eHub                  := starrStationBasisParameter[wStation].stMKs.stSchnittstellendaten.aEintransporte.Hub[Auftragsdaten.wTransferstationsNr1];
      starrStationBasisParameter[wStation].pAuftrag[wWand].stAuftragsOptionen.eHub_NachEintransport := starrStationBasisParameter[wStation].stMKs.stSchnittstellendaten.aEintransporte.HubNachEintransport[Auftragsdaten.wTransferstationsNr1];
      starrStationBasisParameter[wStation].pAuftrag[wWand].stAuftragsOptionen.eHub_NachAustransport := 0;
      starrStationBasisParameter[wStation].pAuftrag[wWand].stAuftragsOptionen.eQuerachse := 0;
      starrStationBasisParameter[wStation].pAuftrag[wWand].stAuftragsOptionen.eAchsrichtung := starrStationBasisParameter[wStation].stMKs.stSchnittstellendaten.aEintransporte.Achsrichtung[Auftragsdaten.wTransferstationsNr1];
      starrStationBasisParameter[wStation].pAuftrag[wWand].stAuftragsOptionen.wMaxTransportGeschwindigkeit:= 0;

      IF ( Auftragsdaten.wTransferwand = cWAND_1 ) THEN
        starrStationBasisParameter[wStation].bScheibentrennen[wWand] := NOT Auftragsdaten.stAuftragsInformationen.cBIT_SRC_WALL_1_EMPTY;
      ELSE
        starrStationBasisParameter[wStation].bScheibentrennen[wWand] := NOT Auftragsdaten.stAuftragsInformationen.cBIT_SRC_WALL_2_EMPTY;
      END_IF
      starrStationBasisParameter[wStation].bRueckwaertsTransportieren[wWand] := ( starrStationBasisParameter[wStation].stMKs.stSchnittstellendaten.aEintransporte.Station[Auftragsdaten.wTransferstationsNr1] = Rueckwaertig );

      steplSchritt := STEP_45_E;

    // EINTRANSPORT ==================================================
    STEP_45_E:
      // Im Step 45 wird in dem vererbten FB Anlagenspezifische Auftragsoptionen gesetzt
      starrStationBasisParameter[wStation].bEintransport[wWand] := TRUE;
      steplSchritt := STEP_50_E;

    // EINTRANSPORT ==================================================
    STEP_50_E:
      (* Hinweis:
         - Scheibenzaehler dekrementieren
         - Scheibe quittieren, sofern dies nötig ist
      *)
      blStationQuittiertScheiben := starrStationBasisParameter[wStation].stMKs.stSchnittstellendaten.aEintransporte.bStationQuittiertScheibe[wlEintransportstation];

      IF ( starrStationBasisParameter[wStation].OutGlasTransport[wWand].bQuittScheibe ) THEN

        IF ( ilScheibenZuQuittieren > 0 ) AND blStationQuittiertScheiben THEN

          wSps2MmiZielStation  := starrStationBasisParameter[wStation].stMKs.stStationsNummern.NummerIntern;
          wSps2MmiQuellStation := Auftragsdaten.wTransferstationsNr1;
          wSps2MmiZielWand     := Auftragsdaten.wStationsWand;
          wSps2MmiQuellWand    := Auftragsdaten.wTransferwand;
          dwSps2MmiWartezeit   := starrStationBasisParameter[wStation].dwWartezeit[wWand];
          wSPS2MMIAuftragstyp  := 0;

          MsgToMmi(auftragsnr_w := SB0_SPS_QUIT_SHEET_ORDER );

        END_IF

        ilScheibenZuQuittieren := ilScheibenZuQuittieren - 1;

      END_IF

      (* Hinweis:
         - Abschliessen des Eintransports
      *)
      IF ( starrStationBasisParameter[wStation].bEintransportAbgeschlossen[wWand] ) THEN
        starrStationBasisParameter[wStation].bRueckwaertsTransportieren[wWand] := FALSE;
        starrStationBasisParameter[wStation].bEintransport[wWand] := FALSE;
        steplSchritt := STEP_1000_E;
      END_IF

      (* Fehlerbehandlung:
         - Station
      *)
      IF ( starrStationBasisParameter[wStation].bFehler ) THEN
        SpsError( eFehler_Station,
                  starrStationBasisParameter[wStation].wFehlerNummer,
                  starrStationBasisParameter[wStation].stMKs.stStationsNummern.NummerIntern,
                  AutomatikkreisBestimmen(starrStationBasisParameter[wStation].stMKs.stStationsNummern.NummerSPS),
                  starrStationBasisParameter[wStation].awFehlerInformationen );

        starrStationBasisParameter[wStation].bEintransport[wWand] := FALSE;
        starrStationBasisParameter[wStation].bRueckwaertsTransportieren[wWand] := FALSE;
        steplSchritt := STEP_900_E;
      END_IF

    // EINTRANSPORT ==================================================
    STEP_100_E:
      // ---------------------------------------------------------------------------------------
      //  OPTIONAL - PRUEFUNG DER SCHEIBENQUITTIERUNG
      //
      //  Hinweis:
      // - n/c
      // ---------------------------------------------------------------------------------------

      IF ( ilScheibenZuQuittieren = 0) THEN
        steplSchritt := STEP_1000_E;

      (* Anmerkung:
         - Zu wenig Scheiben quittiert
      *)
      ELSIF ( ilScheibenZuQuittieren > 0 ) THEN
        wpgFehlerdaten[0] := starrStationBasisParameter[wStation].stMKs.stStationsNummern.NummerExtern;
        wpgFehlerdaten[1] := wWand;
        SpsError( eFehler_Station,
                  cMELDUNG_STATION_ZUWENIG_SCHEIBEN_QUITTIERT_EINTRANSPORT,
                  starrStationBasisParameter[wStation].stMKs.stStationsNummern.NummerIntern,
                  AutomatikkreisBestimmen(starrStationBasisParameter[wStation].stMKs.stStationsNummern.NummerSPS),
                  wpgFehlerdaten );
        steplSchritt := STEP_900_E;

      (* Anmerkung:
         - Zu viele Scheiben quittiert
      *)
      ELSIF ( ilScheibenZuQuittieren < 0 ) THEN
        wpgFehlerdaten[0] := starrStationBasisParameter[wStation].stMKs.stStationsNummern.NummerExtern;
        wpgFehlerdaten[1] := wWand;
        SpsError( eFehler_Station,
                  cMELDUNG_STATION_ZUVIELE_SCHEIBEN_QUITTIERT_EINTRANSPORT,
                  starrStationBasisParameter[wStation].stMKs.stStationsNummern.NummerIntern,
                  AutomatikkreisBestimmen(starrStationBasisParameter[wStation].stMKs.stStationsNummern.NummerSPS),
                  wpgFehlerdaten );
        steplSchritt := STEP_900_E;

      END_IF

    // EINTRANSPORT ==================================================
    STEP_900_E:
      bpFehler := TRUE;

    // EINTRANSPORT ==================================================
    STEP_1000_E:
      bpDone := TRUE;
      IF starrStationBasisParameter[wStation].stMKs.stStationsOptionen.bScheibeAbnehmenNachEintransport THEN
        Auftragsdaten.wAuftrag := eStation_Abnehmen;
      ELSIF Auftragsdaten.bLetzteScheibe THEN
        Auftragsdaten.wAuftrag := eStation_Warte_Auf_Austransport;
      ELSE
        Auftragsdaten.wAuftrag := eStation_Belegt;
      END_IF

  // EINTRANSPORT ==================================================
  END_CASE
END_IF

IF bpReset THEN
  bpFehler := FALSE;
  bpReset := FALSE;
  bpDone := FALSE;
  steplSchritt := STEP_0_E;
  starrStationBasisParameter[wStation].bScheibentrennen[wWand] := FALSE;
  starrStationBasisParameter[wStation].bRueckwaertsTransportieren[wWand] := FALSE;
  starrStationBasisParameter[wStation].bEintransport[wWand] := FALSE;
END_IF
END_FUNCTION_BLOCK

(* ---- Station_Glashoehenmessung.fb.st ---- *)
(* METADATA
{
	"v3Meta": {
		"objectGuid": "4b81b4a3-bc49-4a0d-8ff1-d84de9c8f53e"
	}
}
*)
FUNCTION_BLOCK Station_Glashoehenmessung
VAR_INPUT

  // BOOLEAN
  bpReset                : BOOL;
  bpAbbruchAnlegeauftrag : BOOL;

  // WORD
  wStation               : WORD;

  // STRUKTUR
  Auftragsdaten          : Auftragsdaten_ST;

END_VAR
VAR_OUTPUT

  // BOOLEAN
  bpDone                 : BOOL;
  bpFehler               : BOOL;

END_VAR
VAR

  // STEPS
  steplSchritt           : STEPS_TE;

END_VAR
//-------------------------------------------------------------------------------------------------
// STEUERUNG ANLEGEN
//-------------------------------------------------------------------------------------------------
IF ( Auftragsdaten.wAuftrag = eStation_Hoehenmessung ) THEN
  CASE steplSchritt OF
    // HÖHENMESSUNG ==================================================
    STEP_0_E:
      (* Hinweis:
         - Ueberpruefung des Sicherheitskreises
      *)
      IF checkSafetyCircuitsNotBlocked(starrStationBasisParameter[wStation], eSKKomponente_Messachse) THEN
        steplSchritt := STEP_10_E;
      END_IF

      (* Hinweis:
         - Abbruch des Anlegens
      *)
      IF ( bpAbbruchAnlegeauftrag ) THEN
        bpAbbruchAnlegeauftrag := FALSE;
        bpDone := TRUE;
        Auftragsdaten.wAuftrag := eStation_Kein_Auftrag;
      END_IF

    // HÖHENMESSUNG ==================================================
    STEP_10_E:
      (* Hinweis:
         - Starten des Messvorgangs
      *)
      starrStationBasisParameter[wStation].pAuftrag[cWAND_1] := Auftragsdaten;
      starrStationBasisParameter[wStation].bGlashoehenmessung := TRUE;

      steplSchritt := STEP_20_E;

    // HÖHENMESSUNG ==================================================
    STEP_20_E:
      (* Hinweis:
         - Prüfen dass der Auftragsstatus sich geändert hat
      *)
      IF ( starrStationBasisParameter[wStation].eStatusAuftrag = eAuftragAktiv ) THEN
        steplSchritt := STEP_100_E;
      END_IF

      (* Fehlerbehandlung:
         - Station
      *)
      IF ( starrStationBasisParameter[wStation].bFehler ) THEN
        SpsError( eFehler_Station,
                  starrStationBasisParameter[wStation].wFehlerNummer,
                  starrStationBasisParameter[wStation].stMKs.stStationsNummern.NummerIntern,
                  AutomatikkreisBestimmen(starrStationBasisParameter[wStation].stMKs.stStationsNummern.NummerSPS),
                  starrStationBasisParameter[wStation].awFehlerInformationen );
        starrStationBasisParameter[wStation].bGlashoehenmessung := FALSE;
        steplSchritt := STEP_900_E;
      END_IF

    // HÖHENMESSUNG ==================================================
    STEP_100_E:
      (* Hinweis:
         - Starten des Messvorgangs
      *)
      IF ( starrStationBasisParameter[wStation].bGlashoehenmessungAbgeschlossen ) THEN
        starrStationBasisParameter[wStation].bGlashoehenmessung := FALSE;

        steplSchritt := STEP_1000_E;
      END_IF

      (* Fehlerbehandlung:
         - Station
      *)
      IF ( starrStationBasisParameter[wStation].bFehler ) THEN
        SpsError( eFehler_Station,
                  starrStationBasisParameter[wStation].wFehlerNummer,
                  starrStationBasisParameter[wStation].stMKs.stStationsNummern.NummerIntern,
                  AutomatikkreisBestimmen(starrStationBasisParameter[wStation].stMKs.stStationsNummern.NummerSPS),
                  starrStationBasisParameter[wStation].awFehlerInformationen );

        starrStationBasisParameter[wStation].bGlashoehenmessung := FALSE;
        steplSchritt := STEP_900_E;
      END_IF

    // HÖHENMESSUNG ==================================================
    STEP_900_E:
      bpFehler := TRUE;

    // HÖHENMESSUNG ==================================================
    STEP_1000_E:
      (* Hinweis:
         - Entsprechend dem Auftragsergebnis den Folgeauftrag zuweisen
      *)
      bpDone := TRUE;

      IF ( starrStationBasisParameter[wStation].eStatusAuftrag = eAuftragErfolgreich ) THEN
        Auftragsdaten.wAuftrag := eStation_Messfahrt;

      ELSIF ( starrStationBasisParameter[wStation].eStatusAuftrag = eAuftragWiederholen ) THEN
        Auftragsdaten.wAuftrag := eStation_Anlegen;

      END_IF

  // HÖHENMESSUNG ==================================================
  END_CASE
END_IF

IF bpReset THEN
  bpFehler := FALSE;
  bpReset := FALSE;
  bpDone := FALSE;
  steplSchritt := STEP_0_E;
  starrStationBasisParameter[wStation].bGlashoehenmessung := FALSE;
END_IF
END_FUNCTION_BLOCK

(* ---- Station_Glaslaengenmessung.fb.st ---- *)
(* METADATA
{
	"v3Meta": {
		"objectGuid": "379bb71f-09e3-4346-a24a-24b89454f93a"
	}
}
*)
FUNCTION_BLOCK Station_Glaslaengenmessung
VAR_INPUT

  // BOOLEAN
  bpReset                : BOOL;
  bpAbbruchAnlegeauftrag : BOOL;

  // WORD
  wStation               : WORD;

  // STRUKTUR
  Auftragsdaten          : Auftragsdaten_ST;

END_VAR
VAR_OUTPUT

  // BOOLEAN
  bpDone                 : BOOL;
  bpFehler               : BOOL;

END_VAR
VAR

  // STEPS
  steplSchritt           : STEPS_TE;

END_VAR
//-------------------------------------------------------------------------------------------------
// STEUERUNG: MESSUNG
//-------------------------------------------------------------------------------------------------
IF ( Auftragsdaten.wAuftrag = eStation_Messfahrt ) THEN
  CASE steplSchritt OF
    // MESSFAHRT ==================================================
    STEP_0_E:
      (* Hinweis:
         - Ueberpruefung des Sicherheitskreises
      *)
      IF checkSafetyCircuitsNotBlocked(starrStationBasisParameter[wStation], eSKKomponente_Glastransport) THEN
        steplSchritt := STEP_10_E;
      END_IF

      (* Hinweis:
         - Abbruch des Anl
      *)
      IF ( bpAbbruchAnlegeauftrag ) THEN
        bpAbbruchAnlegeauftrag := FALSE;
        bpDone := TRUE;
        Auftragsdaten.wAuftrag := eStation_Kein_Auftrag;
      END_IF

    // MESSFAHRT ==================================================
    STEP_10_E:
      // Glastyp festlegen
      IF ( Auftragsdaten.rAuftragsLaenge > ( starrStationBasisParameter[wStation].stParameterStationskomponenten.stGlastransport[1].rMessstrecke - rgMKWegAnlegetischUebergroesseScheibeBerechnen ) ) THEN
        starrStationBasisParameter[wStation].wGlasTyp[cWAND_1] := eScheibe_Maximal;
      ELSE
        starrStationBasisParameter[wStation].wGlasTyp[cWAND_1] := eScheibe_Default;
      END_IF

      steplSchritt := STEP_20_E;

    // MESSFAHRT ==================================================
    STEP_20_E:
      (* Hinweis:
         - cMittlereScheibe
           cGrosseScheibe:
           => 1. Option: Anlegetisch kann die Glasvermessung starten ohne die Nachfolgestation
         - cMaxScheibe:
           => 1. Option: Zum vermessen der Scheibe wird die Nachfolgestation benoetigt
      *)
      CASE starrStationBasisParameter[wStation].wGlasTyp[cWAND_1] OF

        cMAXSCHEIBE:
          IF ( Job_Stationen.AuftragsdatenWand[starrStationBasisParameter[wStation].stMKs.stSchnittstellendaten.wNachfolgerStation, cWAND_1].wAuftrag = eStation_Kein_Auftrag ) THEN
            Job_Stationen.AuftragsdatenWand[starrStationBasisParameter[wStation].stMKs.stSchnittstellendaten.wNachfolgerStation, cWAND_1]          := AuftragsdatenUmkopieren(FALSE, FALSE, Auftragsdaten);
            Job_Stationen.AuftragsdatenWand[starrStationBasisParameter[wStation].stMKs.stSchnittstellendaten.wNachfolgerStation, cWAND_1].wAuftrag := eStation_Messkopplung;

            steplSchritt := STEP_30_E;
          END_IF

        ELSE
          steplSchritt := STEP_30_E;

      END_CASE

    // MESSFAHRT ==================================================
    STEP_30_E:
      (* Hinweis:
         - Auftragsdaten uebergeben
         - Starten der Glasmessung
      *)
      starrStationBasisParameter[wStation].pAuftrag[cWAND_1] := Auftragsdaten;
      starrStationBasisParameter[wStation].bGlaslaengenmessung := TRUE;

      steplSchritt := STEP_40_E;

    // MESSFAHRT ==================================================
    STEP_40_E:
      (* Hinweis:
         - Prüfen dass der Auftragsstatus sich geändert hat
      *)
      IF ( starrStationBasisParameter[wStation].eStatusAuftrag = eAuftragAktiv ) THEN
        steplSchritt := STEP_100_E;
      END_IF

    // MESSFAHRT ==================================================
    STEP_100_E:
      (* Hinweis:
         - Glasvermessung abgeschlossen
           => Scheibenvermessung war erfolgreich [Wechsel in den Austransport]
      *)
      IF ( starrStationBasisParameter[wStation].bGlaslaengenmessungAbgeschlossen ) THEN
        starrStationBasisParameter[wStation].bGlaslaengenmessung := FALSE;

        (* Hinweis:
           - Pruefen ob die Betriebsart wieder zurueckgesetzt werden muss
        *)
        steplSchritt := STEP_800_E;

      END_IF

      (* Fehlerbehandlung:
         - Anlegetisch
      *)
      IF ( starrStationBasisParameter[wStation].bFehler ) THEN
        SpsError( eFehler_Station,
                  starrStationBasisParameter[wStation].wFehlerNummer,
                  starrStationBasisParameter[wStation].stMKs.stStationsNummern.NummerIntern,
                  AutomatikkreisBestimmen(starrStationBasisParameter[wStation].stMKs.stStationsNummern.NummerSPS),
                  starrStationBasisParameter[wStation].awFehlerInformationen );

        starrStationBasisParameter[wStation].bGlaslaengenmessung := FALSE;
        steplSchritt := STEP_900_E;
      END_IF

    // MESSFAHRT ==================================================
    STEP_800_E:
      (* Hinweis:
         - Ergebnis der Messung prüfen
      *)
      IF ( starrStationBasisParameter[wStation].eStatusAuftrag = eAuftragErfolgreich ) THEN

        wSps2MmiInputtableNummer := starrStationBasisParameter[wStation].stMKs.stStationsNummern.NummerIntern;
        dwSps2MmiWartezeit       := starrStationBasisParameter[wStation].dwWartezeit[cWAND_1];
        MsgToMmi(auftragsnr_w    := SB0_SPS_SortierungQuittInputInQueue);  // Auftrag für den Anlegetisch

        CASE starrStationBasisParameter[wStation].wGlasTyp[cWAND_1] OF

          cMAXSCHEIBE:
            Job_Stationen.abpResetTransportkopplung[starrStationBasisParameter[wStation].stMKs.stSchnittstellendaten.wNachfolgerStation, cWAND_1]  := TRUE;
            Job_Stationen.AuftragsdatenWand[starrStationBasisParameter[wStation].stMKs.stSchnittstellendaten.wNachfolgerStation, cWAND_1].wAuftrag := eStation_Kein_Auftrag;

        END_CASE

        steplSchritt := STEP_1000_E;

      ELSIF ( starrStationBasisParameter[wStation].eStatusAuftrag = eAuftragWiederholen ) THEN

        CASE starrStationBasisParameter[wStation].wGlasTyp[cWAND_1] OF

          cMAXSCHEIBE:
            Job_Stationen.abpResetTransportkopplung[starrStationBasisParameter[wStation].stMKs.stSchnittstellendaten.wNachfolgerStation, cWAND_1] := TRUE;
            Job_Stationen.AuftragsdatenWand[starrStationBasisParameter[wStation].stMKs.stSchnittstellendaten.wNachfolgerStation, cWAND_1].wAuftrag := eStation_Kein_Auftrag;

        END_CASE

        bpDone := TRUE;
        Auftragsdaten.wAuftrag := eStation_Anlegen;

      END_IF

    // MESSFAHRT ==================================================
    STEP_900_E:
      bpFehler := TRUE;

    // MESSFAHRT ==================================================
    STEP_1000_E:
      (* Wichtig:
         - Auftragsstatus zuweisen
      *)
      bpDone := TRUE;

      Auftragsdaten.wAuftrag := eStation_Warte_Auf_Austransport;

  // MESSFAHRT ==================================================
  END_CASE
END_IF

IF bpReset THEN
  bpFehler := FALSE;
  bpReset := FALSE;
  bpDone := FALSE;
  starrStationBasisParameter[wStation].bGlaslaengenmessung := FALSE;
  steplSchritt := STEP_0_E;
END_IF
END_FUNCTION_BLOCK

(* ---- Station_Messkopplung.fb.st ---- *)
(* METADATA
{
	"v3Meta": {
		"objectGuid": "d07d57e1-6a50-4547-ad5d-dd99acc1a5ad"
	}
}
*)
FUNCTION_BLOCK Station_Messkopplung
VAR_INPUT

  // BOOLEAN
  bpReset                : BOOL;

  // WORD
  wStation               : WORD;
  wWand                  : WORD;

  // STRUKTUR
  Auftragsdaten          : Auftragsdaten_ST;

END_VAR
VAR_OUTPUT

  // BOOLEAN
  bpDone                 : BOOL;
  bpFehler               : BOOL;

END_VAR
VAR

  // STEPS
  steplSchritt           : STEPS_TE;

END_VAR
//-------------------------------------------------------------------------------------------------
// STEUERUNG: MESSUNG
//-------------------------------------------------------------------------------------------------
IF ( Auftragsdaten.wAuftrag = eStation_Messkopplung ) THEN
  CASE steplSchritt OF
    // MESSFAHRT ==================================================
    STEP_0_E:
      (* Hinweis:
         - Ueberpruefung des Sicherheitskreises
      *)
      IF checkSafetyCircuitsNotBlocked(starrStationBasisParameter[wStation], eSKKomponente_Glastransport) THEN
        steplSchritt := STEP_30_E;
      END_IF

    // MESSFAHRT ==================================================
    STEP_30_E:
      (* Hinweis:
         - Auftragsdaten uebergeben
         - Starten der Glasmessung
      *)
      starrStationBasisParameter[wStation].pAuftrag[wWand] := Auftragsdaten;

      starrStationBasisParameter[wStation].pAuftrag[wWand].stAuftragsOptionen.eKippen_SollPosition := starrStationBasisParameter[wStation].stMKs.stSchnittstellendaten.aEintransporte.Kippen[starrStationBasisParameter[wStation].stMKs.stSchnittstellendaten.wVorgaengerStation];
      starrStationBasisParameter[wStation].pAuftrag[wWand].stAuftragsOptionen.eHub                 := starrStationBasisParameter[wStation].stMKs.stSchnittstellendaten.aEintransporte.Hub[starrStationBasisParameter[wStation].stMKs.stSchnittstellendaten.wVorgaengerStation];

      IF ( Auftragsdaten.rAuftragsDicke < wgMKScheibenDicke13mm ) THEN
        starrStationBasisParameter[wStation].pAuftrag[wWand].stAuftragsOptionen.eDickenverstellung := eZylinderStellung16mm;
      ELSIF ( Auftragsdaten.rAuftragsDicke <= wgMKScheibenDicke19mm ) THEN
        starrStationBasisParameter[wStation].pAuftrag[wWand].stAuftragsOptionen.eDickenverstellung := eZylinderStellung23mm;
      ELSE
        starrStationBasisParameter[wStation].pAuftrag[wWand].stAuftragsOptionen.eDickenverstellung := eZylinderStellung29mm;
      END_IF

      starrStationBasisParameter[wStation].bMesskopplung[wWand] := TRUE;

      steplSchritt := STEP_100_E;

    // MESSFAHRT ==================================================
    STEP_100_E:
      (* Fehlerbehandlung:
         - Messkopplung
      *)
      IF ( starrStationBasisParameter[wStation].bFehler ) THEN
        SpsError( eFehler_Station,
                  starrStationBasisParameter[wStation].wFehlerNummer,
                  starrStationBasisParameter[wStation].stMKs.stStationsNummern.NummerIntern,
                  AutomatikkreisBestimmen(starrStationBasisParameter[wStation].stMKs.stStationsNummern.NummerSPS),
                  starrStationBasisParameter[wStation].awFehlerInformationen );

        starrStationBasisParameter[wStation].bMesskopplung[wWand] := FALSE;
        steplSchritt := STEP_900_E;
      END_IF

    // MESSFAHRT ==================================================
    STEP_900_E:
      bpFehler := TRUE;

    // MESSFAHRT ==================================================
    STEP_1000_E:
      (* Wichtig:
         - Auftragsstatus zuweisen
      *)
      bpDone := TRUE;

  // MESSFAHRT ==================================================
  END_CASE
END_IF

IF bpReset THEN
  bpFehler := FALSE;
  bpReset := FALSE;
  bpDone := FALSE;
  starrStationBasisParameter[wStation].bMesskopplung[wWand] := FALSE;
  steplSchritt := STEP_0_E;
END_IF
END_FUNCTION_BLOCK

(* ---- Station_Querfahrt.fb.st ---- *)
(* METADATA
{
	"v3Meta": {
		"objectGuid": "54d45b69-8d91-483b-a87f-7b1de952ab2e"
	}
}
*)
FUNCTION_BLOCK Station_Querfahrt
VAR_INPUT

  // BOOLEAN
  bpReset                : BOOL;

  // WORD
  wStation               : WORD;

  // STRUKTUR
  Auftragsdaten          : Auftragsdaten_ST;

END_VAR
VAR_OUTPUT

  // BOOLEAN
  bpDone                 : BOOL;
  bpFehler               : BOOL;

END_VAR
VAR

  // STEPS
  steplSchritt           : STEPS_TE;

  // BAUSTEINE
  PositionierAuftragsdatenPruefen : PositionierAuftragsdatenPruefen;

END_VAR
// ****************************************************9*********************************************
// STEUERUNG: POSITIONIEREN
// *************************************************************************************************

IF ( Auftragsdaten.wAuftrag = eStation_Vorabpositionierung ) THEN
  CASE steplSchritt OF
    // POSITIONIERUNG ===========================================
    STEP_0_E:
      (* Hinweis:
         - Ueberpruefung des Sicherheitskreises
      *)
      IF checkSafetyCircuitsNotBlocked(starrStationBasisParameter[wStation], eSKKomponente_Querfahrt) THEN

        IF ( ABS( starrStationBasisParameter[wStation].rAktuellePositionQuerfahrt - Auftragsdaten.rVorabPosition ) <= rgMKZielPositionToleranz ) THEN
          steplSchritt := STEP_500_E;
        ELSE
          steplSchritt := STEP_5_E;
        END_IF

      END_IF

    // POSITIONIERUNG ===========================================
    STEP_5_E:
      (* Hinweis:
         - Auftragsdaten pruefen
           => Version der Verfahrlogik beachten
      *)
      steplSchritt := STEP_10_E;

      PositionierAuftragsdatenPruefen.rpSollPosition   := Auftragsdaten.rVorabPosition;
      PositionierAuftragsdatenPruefen.wpStationsNummer := wStation;

      PositionierAuftragsdatenPruefen();

      IF ( NOT PositionierAuftragsdatenPruefen.bpErgebnis ) THEN
        steplSchritt := STEP_900_E;
      END_IF

    // POSITIONIERUNG ===========================================
    STEP_10_E:
      (* Hinweis:
         - Uebergabe der Auftragsdaten
      *)
      starrStationBasisParameter[wStation].pAuftragVorabPositionierung := Auftragsdaten;
      starrStationBasisParameter[wStation].bVorabpositionieren := TRUE;

      steplSchritt := STEP_20_E;

    // POSITIONIERUNG ===========================================
    STEP_20_E:
      (* Hinweis:
         - Nachricht absetzen
      *)
      IF ( starrStationBasisParameter[wStation].bUpdateVorabPositionieren = TRUE ) THEN

        wSps2MmiQuittVorabShuttleNr := starrStationBasisParameter[wStation].stMKs.stStationsNummern.NummerIntern;
        rgSPS2MMIExtractionShuttlePosition := starrStationBasisParameter[wStation].rAktuellePositionQuerfahrt;
        MsgToMmi(auftragsnr_w := SB0_SPS_SHUTTLEVORABPOSITIONIERUNGUPDATE );// Quit 2 MMI Scheibe vorne

        starrStationBasisParameter[wStation].bUpdateVorabPositionieren := FALSE;

        steplSchritt := STEP_100_E;

      END_IF

      (* Fehlerbehandlung:
         - Inputshuttle
      *)
      IF ( starrStationBasisParameter[wStation].bFehler ) THEN

        starrStationBasisParameter[wStation].bVorabpositionieren := FALSE;

        SpsError( eFehler_Station,
                  starrStationBasisParameter[wStation].wFehlerNummer,
                  starrStationBasisParameter[wStation].stMKs.stStationsNummern.NummerIntern,
                  AutomatikkreisBestimmen(starrStationBasisParameter[wStation].stMKs.stStationsNummern.NummerSPS),
                  starrStationBasisParameter[wStation].awFehlerInformationen );

        steplSchritt := STEP_900_E;
      END_IF

    // POSITIONIERUNG ===========================================
    STEP_100_E:
      (* Hinweis:
         - Positionierung abgeschlossen
           => Nachricht absetzen
      *)
      IF ( starrStationBasisParameter[wStation].bVorabpositionierenAbgeschlossen ) THEN

        starrStationBasisParameter[wStation].bVorabpositionieren := FALSE;

        wSps2MmiQuittVorabShuttleNr        := starrStationBasisParameter[wStation].stMKs.stStationsNummern.NummerIntern;
        rgSPS2MMIExtractionShuttlePosition := starrStationBasisParameter[wStation].rAktuellePositionQuerfahrt;
        MsgToMmi(auftragsnr_w := SB0_SPS_QUITTSHUTTLEVORABPOSITIONIERUNG );

        steplSchritt := STEP_1000_E;

      END_IF

      (* Fehlerbehandlung:
         - Inputshuttle
      *)
      IF ( starrStationBasisParameter[wStation].bFehler ) THEN
        starrStationBasisParameter[wStation].bVorabpositionieren := FALSE;

        SpsError( eFehler_Station,
                  starrStationBasisParameter[wStation].wFehlerNummer,
                  starrStationBasisParameter[wStation].stMKs.stStationsNummern.NummerIntern,
                  AutomatikkreisBestimmen(starrStationBasisParameter[wStation].stMKs.stStationsNummern.NummerSPS),
                  starrStationBasisParameter[wStation].awFehlerInformationen );

        steplSchritt := STEP_900_E;
      END_IF

    // POSITIONIERUNG ===========================================
    STEP_500_E:
      wSps2MmiQuittVorabShuttleNr := starrStationBasisParameter[wStation].stMKs.stStationsNummern.NummerIntern;
      rgSPS2MMIExtractionShuttlePosition := starrStationBasisParameter[wStation].rAktuellePositionQuerfahrt;
      MsgToMmi(auftragsnr_w := SB0_SPS_SHUTTLEVORABPOSITIONIERUNGUPDATE );
      steplSchritt := STEP_510_E;

    // POSITIONIERUNG ===========================================
    STEP_510_E:
      wSps2MmiQuittVorabShuttleNr        := starrStationBasisParameter[wStation].stMKs.stStationsNummern.NummerIntern;
      rgSPS2MMIExtractionShuttlePosition := starrStationBasisParameter[wStation].rAktuellePositionQuerfahrt;
      MsgToMmi(auftragsnr_w := SB0_SPS_QUITTSHUTTLEVORABPOSITIONIERUNG );
      steplSchritt := STEP_1000_E;

    // POSITIONIERUNG ===========================================
    STEP_900_E:
      bpFehler := TRUE;

    // POSITIONIERUNG ===========================================
    STEP_1000_E:
      bpDone := TRUE;
      Auftragsdaten.wAuftrag := eStation_Kein_Auftrag;

  // POSITIONIERUNG ===========================================
  END_CASE
END_IF

IF bpReset THEN
  bpFehler := FALSE;
  bpDone   := FALSE;
  bpReset  := FALSE;
  Auftragsdaten.wAuftrag := eStation_Kein_Auftrag;
  starrStationBasisParameter[wStation].bUpdateVorabPositionieren := FALSE;
  starrStationBasisParameter[wStation].bVorabpositionieren := FALSE;
  steplSchritt := STEP_0_E;
END_IF
END_FUNCTION_BLOCK

(* ---- Station_Transportkopplung.fb.st ---- *)
(* METADATA
{
	"v3Meta": {
		"objectGuid": "7029972e-eb09-4666-92ad-77d763ae2960"
	}
}
*)
FUNCTION_BLOCK Station_Transportkopplung
VAR_INPUT

  // BOOLEAN
  bpReset                : BOOL;

  // WORD
  wStation               : WORD;
  wWand                  : WORD;

  // STRUKTUR
  Auftragsdaten          : Auftragsdaten_ST;

END_VAR
VAR_OUTPUT

  // BOOLEAN
  bpDone                 : BOOL;
  bpFehler               : BOOL;

END_VAR
VAR

  // STEPS
  steplSchritt           : STEPS_TE;

END_VAR
//-------------------------------------------------------------------------------------------------
// STEUERUNG: MESSUNG
//-------------------------------------------------------------------------------------------------
IF ( Auftragsdaten.wAuftrag = eStation_Transportkopplung ) THEN
  CASE steplSchritt OF
    // MESSFAHRT ==================================================
    STEP_0_E:
      (* Hinweis:
         - Ueberpruefung des Sicherheitskreises
      *)
      IF checkSafetyCircuitsNotBlocked(starrStationBasisParameter[wStation], eSKKomponente_Glastransport) THEN
        steplSchritt := STEP_30_E;
      END_IF

    // MESSFAHRT ==================================================
    STEP_30_E:
      (* Hinweis:
         - Auftragsdaten uebergeben
         - Starten der Glasmessung
      *)
      starrStationBasisParameter[wStation].pAuftrag[wWand] := Auftragsdaten;

      starrStationBasisParameter[wStation].pAuftrag[wWand].stAuftragsOptionen.eKippen_SollPosition := starrStationBasisParameter[wStation].stMKs.stSchnittstellendaten.aEintransporte.Kippen[starrStationBasisParameter[wStation].stMKs.stSchnittstellendaten.wVorgaengerStation];
      starrStationBasisParameter[wStation].pAuftrag[wWand].stAuftragsOptionen.eHub                 := starrStationBasisParameter[wStation].stMKs.stSchnittstellendaten.aEintransporte.Hub[starrStationBasisParameter[wStation].stMKs.stSchnittstellendaten.wVorgaengerStation];

      IF ( Auftragsdaten.rAuftragsDicke < wgMKScheibenDicke13mm ) THEN
        starrStationBasisParameter[wStation].pAuftrag[wWand].stAuftragsOptionen.eDickenverstellung := eZylinderStellung16mm;
      ELSIF ( Auftragsdaten.rAuftragsDicke <= wgMKScheibenDicke19mm ) THEN
        starrStationBasisParameter[wStation].pAuftrag[wWand].stAuftragsOptionen.eDickenverstellung := eZylinderStellung23mm;
      ELSE
        starrStationBasisParameter[wStation].pAuftrag[wWand].stAuftragsOptionen.eDickenverstellung := eZylinderStellung29mm;
      END_IF

      starrStationBasisParameter[wStation].bTransportkopplung[wWand] := TRUE;

      steplSchritt := STEP_100_E;

    // MESSFAHRT ==================================================
    STEP_100_E:
      (* Fehlerbehandlung:
         - Transportkopplung
      *)
      IF ( starrStationBasisParameter[wStation].bFehler ) THEN
        SpsError( eFehler_Station,
                  starrStationBasisParameter[wStation].wFehlerNummer,
                  starrStationBasisParameter[wStation].stMKs.stStationsNummern.NummerIntern,
                  AutomatikkreisBestimmen(starrStationBasisParameter[wStation].stMKs.stStationsNummern.NummerSPS),
                  starrStationBasisParameter[wStation].awFehlerInformationen );

        starrStationBasisParameter[wStation].bTransportkopplung[wWand] := FALSE;
        steplSchritt := STEP_900_E;
      END_IF

    // MESSFAHRT ==================================================
    STEP_900_E:
      bpFehler := TRUE;

    // MESSFAHRT ==================================================
    STEP_1000_E:
      (* Wichtig:
         - Auftragsstatus zuweisen
      *)
      bpDone := TRUE;

  // MESSFAHRT ==================================================
  END_CASE
END_IF

IF bpReset THEN
  bpFehler := FALSE;
  bpReset := FALSE;
  bpDone := FALSE;
  starrStationBasisParameter[wStation].bTransportkopplung[wWand] := FALSE;
  steplSchritt := STEP_0_E;
END_IF
END_FUNCTION_BLOCK

(* ---- Station_Vortransport.fb.st ---- *)
(* METADATA
{
	"v3Meta": {
		"objectGuid": "9f1ab894-d35e-4a4e-8f77-3236b7a1099b"
	}
}
*)
FUNCTION_BLOCK Station_Vortransport
VAR_INPUT

  // BOOLEAN
  bpReset                : BOOL;

  // WORD
  wStation               : WORD;
  wWand                  : WORD;

  // STRUKTUR
  Auftragsdaten          : Auftragsdaten_ST;

END_VAR
VAR_OUTPUT

  // BOOLEAN
  bpDone                 : BOOL;
  bpFehler               : BOOL;

END_VAR
VAR

  // STEPS
  steplSchritt           : STEPS_TE;

END_VAR
//-------------------------------------------------------------------------------------------------
// STEUERUNG: EINTRANSPORT
//-------------------------------------------------------------------------------------------------
IF ( Auftragsdaten.wAuftrag = eStation_Vortransport ) THEN
  CASE steplSchritt OF
    // EINTRANSPORT ==================================================
    STEP_0_E:
      (* Hinweis:
         - Ueberpruefung des Sicherheitskreises
      *)

      IF checkSafetyCircuitsNotBlocked(starrStationBasisParameter[wStation], eSKKomponente_Glastransport) THEN
        steplSchritt := STEP_10_E;
      END_IF

    // EINTRANSPORT ==================================================
    STEP_10_E:
      (* Hinweis:
         - Vortransport starten
      *)
      (* Hinweis:
         - Auftragsdaten zuweisen
      *)
      starrStationBasisParameter[wStation].pAuftrag[wWand] := Auftragsdaten;

      starrStationBasisParameter[wStation].bVortransport[wWand]    := TRUE;

      steplSchritt := STEP_20_E;

    // EINTRANSPORT ==================================================
    STEP_20_E:
      (* Hinweis:
         - Abschliessen des Eintransports
      *)
      IF ( starrStationBasisParameter[wStation].bVortransportAbgeschlossen[wWand] ) THEN
        starrStationBasisParameter[wStation].bVortransport[wWand] := FALSE;
        steplSchritt := STEP_1000_E;
      END_IF

      (* Fehlerbehandlung:
         - Station
      *)
      IF ( starrStationBasisParameter[wStation].bFehler ) THEN
        SpsError( eFehler_Station,
                  starrStationBasisParameter[wStation].wFehlerNummer,
                  starrStationBasisParameter[wStation].stMKs.stStationsNummern.NummerIntern,
                  AutomatikkreisBestimmen(starrStationBasisParameter[wStation].stMKs.stStationsNummern.NummerSPS),
                  starrStationBasisParameter[wStation].awFehlerInformationen );
        starrStationBasisParameter[wStation].bVortransport[wWand] := FALSE;
        steplSchritt := STEP_900_E;
      END_IF

    // EINTRANSPORT ==================================================
    STEP_900_E:
      bpFehler := TRUE;

    // EINTRANSPORT ==================================================
    STEP_1000_E:
      bpDone := TRUE;
      Auftragsdaten.wAuftrag := eStation_Warte_Auf_Austransport;

  // EINTRANSPORT ==================================================
  END_CASE
END_IF

IF bpReset THEN
  bpFehler := FALSE;
  bpReset := FALSE;
  bpDone := FALSE;
  steplSchritt := STEP_0_E;
  starrStationBasisParameter[wStation].bVortransport[wWand] := FALSE;
END_IF
END_FUNCTION_BLOCK

(* ---- TS_Austransport.fb.st ---- *)
(* METADATA
{
	"v3Meta": {
		"objectGuid": "0f3a9f54-24b3-4180-b764-650377bf6b92"
	}
}
*)
FUNCTION_BLOCK TS_Austransport
VAR_INPUT

  // BOOLEAN
  bpReset                : BOOL;

  // WORD
  wStation               : WORD;

  // STRUKTUR
  Auftragsdaten          : Auftragsdaten_ST;

END_VAR
VAR_OUTPUT

  // BOOLEAN
  bpDone                 : BOOL;
  bpFehler               : BOOL;

END_VAR
VAR
  // BOOLEAN
  blStationQuittiertScheiben : BOOL;

  // WORD
  wlAustransportstation  : WORD;

  // INT
  ilScheibenZuQuittieren : INT;

  // STEPS
  steplSchritt           : STEPS_TE;

END_VAR
//-------------------------------------------------------------------------------------------------
// STEUERUNG: AUSTRANSPORT
//-------------------------------------------------------------------------------------------------
IF ( Auftragsdaten.wAuftrag = eStation_Austransport ) THEN
  CASE steplSchritt OF
    // AUSTRANSPORT  ===========================================
    STEP_0_E:
      (* Hinweis:
         - Sicherheitskreis puefen
         - Austransport aktiv
      *)
      IF ( checkSafetyCircuitsNotBlocked(starrTransferShuttleBasisParameter[wStation])
           AND NOT starrTransfershuttleBasisParameter[wStation].bReset )
      THEN
        steplSchritt := STEP_10_E;
      END_IF

    // AUSTRANSPORT  ===========================================
    STEP_10_E:
      (* Anmerkung:
         - Zielstation abfragen ob diese bereit ist zum Austransport
      *)
      wlAustransportstation := Auftragsdaten.wTransferstationsNr1;
      ilScheibenZuQuittieren := WORD_TO_INT(Auftragsdaten.wAnzahlScheiben);

      starrTransfershuttleBasisParameter[wStation].bRueckwaertsTransportieren[cWAND_1] := FALSE;

      CASE wlAustransportstation OF

        (* Hinweis:
           - Verfahrbahrer Speicher
        *)
        // Fremdanlage Auslauf
        //   - Wie beim Shuttle: Der TS legt den Auftrag der Fremdanlage an, sobald diese frei ist
        cERSTE_FREMDANLAGE_AUSLAUF..cLETZTE_FREMDANLAGE_AUSLAUF:
          IF ( Job_Fremdanlage.AuftragsdatenFremdanlage[wlAustransportstation].wAuftrag = eStation_Kein_Auftrag ) THEN

            // Kopplung zur Fremdanlage herstellen
            starrTransfershuttleBasisParameter[wStation].InGlasTransportNachfolger[cWAND_1] := starrFremdanlageAuslaufStationBasisParameter[wlAustransportstation].OutGlasTransport[cWAND_1];
            starrTransfershuttleBasisParameter[wStation].InGlasTransportVorgaenger[cWAND_1] := starrFremdanlageAuslaufStationBasisParameter[wlAustransportstation].OutGlasTransport[cWAND_1];
            starrFremdanlageAuslaufStationBasisParameter[wlAustransportstation].InGlasTransportVorgaenger[cWAND_1] := starrTransfershuttleBasisParameter[wStation].OutGlasTransport[cWAND_1];

            // Auftragsdaten in die Fremdanlage kopieren
            Job_Fremdanlage.AuftragsdatenFremdanlage[wlAustransportstation]          := AuftragsdatenUmkopieren(FALSE, FALSE, Auftragsdaten);
            Job_Fremdanlage.AuftragsdatenFremdanlage[wlAustransportstation].wAuftrag := eStation_Eintransport;

            steplSchritt := STEP_20_E;
          END_IF

        // Stationen
        //   - Wie beim Shuttle: Der TS legt den Eintransport-Auftrag der Station an
        //   - Durchtransportierende Station behaelt ihren Auftrag
        cERSTE_STATION..cLETZTE_STATION:
          IF (    ( Job_Stationen.AuftragsdatenWand[wlAustransportstation, Auftragsdaten.wTransferwand].wAuftrag = eStation_Kein_Auftrag )
               OR ( Job_Stationen.AuftragsdatenWand[wlAustransportstation, Auftragsdaten.wTransferwand].wAuftrag = eStation_Belegt )
               OR ( Job_Stationen.AuftragsdatenWand[wlAustransportstation, Auftragsdaten.wTransferwand].wAuftrag = eStation_Durchtransport ) )
             AND AutomatikAktiv(wlAustransportstation)
          THEN

            IF NOT ( Job_Stationen.AuftragsdatenWand[wlAustransportstation, Auftragsdaten.wTransferwand].wAuftrag = eStation_Durchtransport ) THEN
              Job_Stationen.AuftragsdatenWand[wlAustransportstation, Auftragsdaten.wTransferwand]          := AuftragsdatenUmkopieren(FALSE, FALSE, Auftragsdaten);
              Job_Stationen.AuftragsdatenWand[wlAustransportstation, Auftragsdaten.wTransferwand].wAuftrag := eStation_Eintransport;
            END_IF

            // Kopplung zur Station herstellen
            starrTransfershuttleBasisParameter[wStation].InGlasTransportNachfolger[cWAND_1] := starrStationBasisParameter[wlAustransportstation].OutGlasTransport[Auftragsdaten.wTransferwand];
            starrTransfershuttleBasisParameter[wStation].InGlasTransportVorgaenger[cWAND_1] := starrStationBasisParameter[wlAustransportstation].OutGlasTransport[Auftragsdaten.wTransferwand];

            steplSchritt := STEP_20_E;
          END_IF

        (* Hinweis:
           - Ruecktransport durch den Speicher beruecksichtigen
        *)
        cERSTES_INPUTSHUTTLE..cLETZTES_INPUTSHUTTLE,
        cERSTES_OUTPUTSHUTTLE..cLETZTES_OUTPUTSHUTTLE:
            IF ( Job_Shuttle.AuftragsdatenWand[wlAustransportstation, Auftragsdaten.wTransferwand].wAuftrag  = eStation_Eintransport ) THEN

              // Kopplung zur Station herstellen
              starrTransfershuttleBasisParameter[wStation].InGlasTransportNachfolger[cWAND_1] := starrShuttleBasisParameter[wlAustransportstation].OutGlasTransport[Auftragsdaten.wTransferwand];
              starrTransfershuttleBasisParameter[wStation].InGlasTransportVorgaenger[cWAND_1] := starrShuttleBasisParameter[wlAustransportstation].OutGlasTransport[Auftragsdaten.wTransferwand];

              steplSchritt := STEP_20_E;
            END_IF

          // Ausnahmesituation:
          //   - Shuttle hat den falschen Auftragsstatus
          IF ( Job_Shuttle.AuftragsdatenWand[wlAustransportstation, Auftragsdaten.wTransferwand].wAuftrag  <> eStation_Eintransport ) THEN
            wpgFehlerdaten[0] := starrTransfershuttleBasisParameter[wStation].stMKs.stStationsNummern.NummerExtern;
            wpgFehlerdaten[1] := wlAustransportstation;
            wpgFehlerdaten[2] := Job_Shuttle.AuftragsdatenWand[wlAustransportstation, Auftragsdaten.wTransferwand].wAuftrag;

            SpsError( eFehler_Station,
                      cMELDUNG_AUFTRAGSDATEN_AUFTRAGSTATUS_GLAS_EMPFAENGER_UNGUELTIG,
                      starrTransfershuttleBasisParameter[wStation].stMKs.stStationsNummern.NummerIntern,
                      AutomatikkreisBestimmen(starrTransfershuttleBasisParameter[wStation].stMKs.stStationsNummern.NummerSPS),
                      wpgFehlerdaten );
            steplSchritt := STEP_900_E;
          END_IF

      END_CASE

      (* Fehlerbehandlung:
         - Shuttle
      *)
      IF ( starrTransfershuttleBasisParameter[wStation].bFehler ) THEN
        SpsError( eFehler_Station,
                  starrTransfershuttleBasisParameter[wStation].wFehlerNummer,
                  starrTransfershuttleBasisParameter[wStation].stMKs.stStationsNummern.NummerIntern,
                  AutomatikkreisBestimmen(starrTransfershuttleBasisParameter[wStation].stMKs.stStationsNummern.NummerSPS),
                  starrTransfershuttleBasisParameter[wStation].awFehlerInformationen );

        steplSchritt := STEP_900_E;
      END_IF

    // AUSTRANSPORT  ===========================================
    STEP_20_E:
      (* Hinweis:
         - Starten des Austransport
      *)
      starrTransfershuttleBasisParameter[wStation].pAuftrag[cWAND_1] := Auftragsdaten;
      starrTransfershuttleBasisParameter[wStation].bAustransport[cWAND_1] := TRUE;
      starrTransfershuttleBasisParameter[wStation].bRueckwaertsTransportieren[cWAND_1] := ( starrTransferShuttleBasisParameter[wStation].stMKs.stSchnittstellendaten.aAustransporte.Station[wlAustransportstation] = Rueckwaertig );
      ilScheibenZuQuittieren := WORD_TO_INT( Auftragsdaten.wAnzahlScheiben);

      steplSchritt := STEP_400_E;

    // AUSTRANSPORT ===============================================
    STEP_400_E:
      // ---------------------------------------------------------------------------------------
      //  QUITTIERUNGEN UND AUSTRANSPORT- ABSCHLUSS
      //
      //  Hinweis:
      //  - Scheibenquittieren: Message zur MMI
      // ---------------------------------------------------------------------------------------

      IF ( starrTransfershuttleBasisParameter[wStation].OutGlasTransport[cWAND_1].bQuittScheibe ) THEN

        IF ( ilScheibenZuQuittieren > 0 ) AND starrTransfershuttleBasisParameter[wStation].stMKs.stSchnittstellendaten.aAustransporte.bStationQuittiertScheibe[wlAustransportstation] THEN

          wSps2MmiZielStation  := Auftragsdaten.wTransferstationsNr1;
          wSps2MmiQuellStation := starrTransfershuttleBasisParameter[wStation].stMKs.stStationsNummern.NummerIntern;
          wSps2MmiZielWand     := Auftragsdaten.wTransferwand;
          wSps2MmiQuellWand    := cWAND_1;
          dwSps2MmiWartezeit   := starrTransfershuttleBasisParameter[wStation].dwWartezeit[cWAND_1];
          wSPS2MMIAuftragstyp  := 1;

          MsgToMmi(auftragsnr_w := SB0_SPS_QUIT_SHEET_ORDER );
        END_IF

        ilScheibenZuQuittieren := ilScheibenZuQuittieren - 1;

      END_IF

      (* Hinweis:
         - Abschliessen des Austransports
      *)
      IF ( starrTransfershuttleBasisParameter[wStation].bAustransportAbgeschlossen[cWAND_1] ) THEN

        starrTransfershuttleBasisParameter[wStation].bAustransport[cWAND_1]                 := FALSE;
        starrTransfershuttleBasisParameter[wStation].bRueckwaertsTransportieren[cWAND_1]    := FALSE;

        steplSchritt := STEP_410_E;
      END_IF

      (* Fehlerbehandlung:
         - Transfershuttle
      *)
      IF ( starrTransfershuttleBasisParameter[wStation].bFehler ) THEN

        IF ( aTransfershuttles[wStation].bpAnforderungBetriebsstopp ) THEN

          (* Hinweis:
             - Ausnahmefehler des TS an die MMI melden
          *)
          IF ( bgAktivierungTransfershuttleSystemcheck ) THEN
            wgSps2MmiShuttleNr                 := starrTransfershuttleBasisParameter[wStation].stMKs.stStationsNummern.NummerIntern;
            wSps2MmiFehlertyp                  := aTransfershuttles[wStation].wpAusnahmefehlerTyp;
            MsgToMmi(auftragsnr_w := SB0_SPS_TRANSFERSHUTTLEFEHLER );
          END_IF

          bpFehler := TRUE;

        END_IF

        starrTransfershuttleBasisParameter[wStation].bAustransport[cWAND_1] := FALSE;
        SpsError( eFehler_Station,
                  starrTransfershuttleBasisParameter[wStation].wFehlerNummer,
                  starrTransfershuttleBasisParameter[wStation].stMKs.stStationsNummern.NummerIntern,
                  AutomatikkreisBestimmen(starrTransfershuttleBasisParameter[wStation].stMKs.stStationsNummern.NummerSPS),
                  starrTransfershuttleBasisParameter[wStation].awFehlerInformationen );

        steplSchritt := STEP_900_E;
      END_IF

    // AUSTRANSPORT ==============================================
    STEP_410_E:
      (* Anmerkung:
         - Gueltige Anzahl von Scheiben wurden quittiert
      *)
      IF ( ilScheibenZuQuittieren = 0 ) THEN
        starrTransfershuttleBasisParameter[wStation].bAustransport[cWAND_1] := FALSE;
        steplSchritt := STEP_1000_E;

      (* Anmerkung:
         - Zu wenig Scheiben quittiert
      *)
      ELSIF ( ilScheibenZuQuittieren > 0 ) THEN
        wpgFehlerdaten[0] := starrTransfershuttleBasisParameter[wStation].stMKs.stStationsNummern.NummerExtern;
        wpgFehlerdaten[1] := cWAND_1;

        SpsError( eFehler_Station,
                  cMELDUNG_STATION_ZUWENIG_SCHEIBEN_QUITTIERT_WAND_AUSTRANSPORT,
                  starrTransfershuttleBasisParameter[wStation].stMKs.stStationsNummern.NummerIntern,
                  AutomatikkreisBestimmen(starrTransfershuttleBasisParameter[wStation].stMKs.stStationsNummern.NummerSPS),
                  wpgFehlerdaten );

        starrTransfershuttleBasisParameter[wStation].bAustransport[cWAND_1] := FALSE;
        steplSchritt := STEP_900_E;

      (* Anmerkung:
         - Zu viele Scheiben quittiert
      *)
      ELSIF ( ilScheibenZuQuittieren < 0 ) THEN
        wpgFehlerdaten[0] := starrTransfershuttleBasisParameter[wStation].stMKs.stStationsNummern.NummerExtern;
        wpgFehlerdaten[1] := cWAND_1;

        SpsError( eFehler_Station,
                  cMELDUNG_STATION_ZUVIELE_SCHEIBEN_QUITTIERT_WAND_AUSTRANSPORT,
                  starrTransfershuttleBasisParameter[wStation].stMKs.stStationsNummern.NummerIntern,
                  AutomatikkreisBestimmen(starrTransfershuttleBasisParameter[wStation].stMKs.stStationsNummern.NummerSPS),
                  wpgFehlerdaten );

        starrTransfershuttleBasisParameter[wStation].bAustransport[cWAND_1] := FALSE;
        steplSchritt := STEP_900_E;
      END_IF

    // AUSTRANSPORT  ===========================================
    STEP_900_E:
      bpFehler := TRUE;

    // AUSTRANSPORT  ===========================================
    STEP_1000_E:
      bpDone := TRUE;

      Auftragsdaten.wAuftrag := eStation_Kein_Auftrag;

      (* Hinweis:
         - Pruefen ob die Transferkopplung geloest werden muss
      *)
      IF ( PruefungWertImIntervall(Auftragsdaten.wTransferstationsNr2, cERSTES_TRANSFERSHUTTLE, cLETZTES_TRANSFERSHUTTLE) ) THEN

        IF ( Job_Shuttle.AuftragsdatenTransfershuttle[Auftragsdaten.wTransferstationsNr2].wAuftrag = eStation_Transportkopplung ) THEN
          Job_Shuttle.abpResetTransportkopplung[Auftragsdaten.wTransferstationsNr2] := TRUE;
        END_IF

      END_IF

  // AUSTRANSPORT  ===========================================
  END_CASE
END_IF

IF bpReset THEN
  bpDone := FALSE;
  bpReset := FALSE;
  bpFehler := FALSE;
  starrTransfershuttleBasisParameter[wStation].bAustransport[cWAND_1] := FALSE;
  steplSchritt := STEP_0_E;
END_IF
END_FUNCTION_BLOCK
